(* IEC 61131-3 sources: 2026_Projet_YGO_ExcavatriceDragage/TOOLS/TEST_AUTO_CI/RESULTS/L_SIMULATION/tests (part 9) *)

TEST 'TC-T418-INT-007 Config maintien reel trop long refuse sans bypass'
nx := 5000; ny := 5000; raw1 := 0; raw2 := 0; previousButton := FALSE; buttonEdges := 0;
bench.Enable := TRUE; joy.Enable := TRUE; joy.ArmingPermit := TRUE; diagOk.Operational := TRUE;
joy.BusCanOpenOP := diagOk; joy.JoystickOP := diagOk; home.Enable := TRUE; home.BootReady := TRUE;
home.Mode := E_Mode.MAINT_N1; home.BucketOffsetValid := TRUE; home.WinchesMechanicallyStopped := TRUE;
cfg.DeadmanArmHoldTime := T#1S;
ADVANCE_TIME(10000000);
bench(RawPosM1 := raw1, RawPosM2 := raw2);
joy(RawX := bench.Operator.JoyXRaw_ANA1, RawY := bench.Operator.JoyYRaw_ANA2, RawButton := bench.Operator.JoyBtnRaw, Cfg := cfg, NeutralXMem := nx, NeutralYMem := ny);
home(DeadmanArmed := joy.DeadmanArmed, JoystickDeflected := NOT joy.AtNeutralXY, JoystickPull := joy.AxisCmdY.DirectionPositive, JoystickPush := joy.AxisCmdY.DirectionNegative, BtnValidation := bench.Operator.JoyBtnRaw);
IF bench.Operator.JoyBtnRaw AND NOT previousButton THEN buttonEdges := buttonEdges + 1; END_IF; previousButton := bench.Operator.JoyBtnRaw;
bench.SimJoystickRight_Fwd_MAINT_Active := TRUE;
ADVANCE_TIME(10000000);
bench(RawPosM1 := raw1, RawPosM2 := raw2);
joy(RawX := bench.Operator.JoyXRaw_ANA1, RawY := bench.Operator.JoyYRaw_ANA2, RawButton := bench.Operator.JoyBtnRaw, Cfg := cfg, NeutralXMem := nx, NeutralYMem := ny);
home(DeadmanArmed := joy.DeadmanArmed, JoystickDeflected := NOT joy.AtNeutralXY, JoystickPull := joy.AxisCmdY.DirectionPositive, JoystickPush := joy.AxisCmdY.DirectionNegative, BtnValidation := bench.Operator.JoyBtnRaw);
IF bench.Operator.JoyBtnRaw AND NOT previousButton THEN buttonEdges := buttonEdges + 1; END_IF; previousButton := bench.Operator.JoyBtnRaw;
ASSERT_FALSE(joy.DeadmanArmed, 'Maintien reel superieur a appui simule donc refus'); ASSERT_FALSE(joy.AxisCmdX.StartStop, 'Aucun bypass');
ADVANCE_TIME(10000000);
bench(RawPosM1 := raw1, RawPosM2 := raw2);
joy(RawX := bench.Operator.JoyXRaw_ANA1, RawY := bench.Operator.JoyYRaw_ANA2, RawButton := bench.Operator.JoyBtnRaw, Cfg := cfg, NeutralXMem := nx, NeutralYMem := ny);
home(DeadmanArmed := joy.DeadmanArmed, JoystickDeflected := NOT joy.AtNeutralXY, JoystickPull := joy.AxisCmdY.DirectionPositive, JoystickPush := joy.AxisCmdY.DirectionNegative, BtnValidation := bench.Operator.JoyBtnRaw);
IF bench.Operator.JoyBtnRaw AND NOT previousButton THEN buttonEdges := buttonEdges + 1; END_IF; previousButton := bench.Operator.JoyBtnRaw;
ASSERT_FALSE(joy.DeadmanArmed, 'Maintien reel superieur a appui simule donc refus'); ASSERT_FALSE(joy.AxisCmdX.StartStop, 'Aucun bypass');
ADVANCE_TIME(10000000);
bench(RawPosM1 := raw1, RawPosM2 := raw2);
joy(RawX := bench.Operator.JoyXRaw_ANA1, RawY := bench.Operator.JoyYRaw_ANA2, RawButton := bench.Operator.JoyBtnRaw, Cfg := cfg, NeutralXMem := nx, NeutralYMem := ny);
home(DeadmanArmed := joy.DeadmanArmed, JoystickDeflected := NOT joy.AtNeutralXY, JoystickPull := joy.AxisCmdY.DirectionPositive, JoystickPush := joy.AxisCmdY.DirectionNegative, BtnValidation := bench.Operator.JoyBtnRaw);
IF bench.Operator.JoyBtnRaw AND NOT previousButton THEN buttonEdges := buttonEdges + 1; END_IF; previousButton := bench.Operator.JoyBtnRaw;
ASSERT_FALSE(joy.DeadmanArmed, 'Maintien reel superieur a appui simule donc refus'); ASSERT_FALSE(joy.AxisCmdX.StartStop, 'Aucun bypass');
ADVANCE_TIME(10000000);
bench(RawPosM1 := raw1, RawPosM2 := raw2);
joy(RawX := bench.Operator.JoyXRaw_ANA1, RawY := bench.Operator.JoyYRaw_ANA2, RawButton := bench.Operator.JoyBtnRaw, Cfg := cfg, NeutralXMem := nx, NeutralYMem := ny);
home(DeadmanArmed := joy.DeadmanArmed, JoystickDeflected := NOT joy.AtNeutralXY, JoystickPull := joy.AxisCmdY.DirectionPositive, JoystickPush := joy.AxisCmdY.DirectionNegative, BtnValidation := bench.Operator.JoyBtnRaw);
IF bench.Operator.JoyBtnRaw AND NOT previousButton THEN buttonEdges := buttonEdges + 1; END_IF; previousButton := bench.Operator.JoyBtnRaw;
ASSERT_FALSE(joy.DeadmanArmed, 'Maintien reel superieur a appui simule donc refus'); ASSERT_FALSE(joy.AxisCmdX.StartStop, 'Aucun bypass');
ADVANCE_TIME(10000000);
bench(RawPosM1 := raw1, RawPosM2 := raw2);
joy(RawX := bench.Operator.JoyXRaw_ANA1, RawY := bench.Operator.JoyYRaw_ANA2, RawButton := bench.Operator.JoyBtnRaw, Cfg := cfg, NeutralXMem := nx, NeutralYMem := ny);
home(DeadmanArmed := joy.DeadmanArmed, JoystickDeflected := NOT joy.AtNeutralXY, JoystickPull := joy.AxisCmdY.DirectionPositive, JoystickPush := joy.AxisCmdY.DirectionNegative, BtnValidation := bench.Operator.JoyBtnRaw);
IF bench.Operator.JoyBtnRaw AND NOT previousButton THEN buttonEdges := buttonEdges + 1; END_IF; previousButton := bench.Operator.JoyBtnRaw;
ASSERT_FALSE(joy.DeadmanArmed, 'Maintien reel superieur a appui simule donc refus'); ASSERT_FALSE(joy.AxisCmdX.StartStop, 'Aucun bypass');
ADVANCE_TIME(10000000);
bench(RawPosM1 := raw1, RawPosM2 := raw2);
joy(RawX := bench.Operator.JoyXRaw_ANA1, RawY := bench.Operator.JoyYRaw_ANA2, RawButton := bench.Operator.JoyBtnRaw, Cfg := cfg, NeutralXMem := nx, NeutralYMem := ny);
home(DeadmanArmed := joy.DeadmanArmed, JoystickDeflected := NOT joy.AtNeutralXY, JoystickPull := joy.AxisCmdY.DirectionPositive, JoystickPush := joy.AxisCmdY.DirectionNegative, BtnValidation := bench.Operator.JoyBtnRaw);
IF bench.Operator.JoyBtnRaw AND NOT previousButton THEN buttonEdges := buttonEdges + 1; END_IF; previousButton := bench.Operator.JoyBtnRaw;
ASSERT_FALSE(joy.DeadmanArmed, 'Maintien reel superieur a appui simule donc refus'); ASSERT_FALSE(joy.AxisCmdX.StartStop, 'Aucun bypass');
ADVANCE_TIME(10000000);
bench(RawPosM1 := raw1, RawPosM2 := raw2);
joy(RawX := bench.Operator.JoyXRaw_ANA1, RawY := bench.Operator.JoyYRaw_ANA2, RawButton := bench.Operator.JoyBtnRaw, Cfg := cfg, NeutralXMem := nx, NeutralYMem := ny);
home(DeadmanArmed := joy.DeadmanArmed, JoystickDeflected := NOT joy.AtNeutralXY, JoystickPull := joy.AxisCmdY.DirectionPositive, JoystickPush := joy.AxisCmdY.DirectionNegative, BtnValidation := bench.Operator.JoyBtnRaw);
IF bench.Operator.JoyBtnRaw AND NOT previousButton THEN buttonEdges := buttonEdges + 1; END_IF; previousButton := bench.Operator.JoyBtnRaw;
ASSERT_FALSE(joy.DeadmanArmed, 'Maintien reel superieur a appui simule donc refus'); ASSERT_FALSE(joy.AxisCmdX.StartStop, 'Aucun bypass');
ADVANCE_TIME(10000000);
bench(RawPosM1 := raw1, RawPosM2 := raw2);
joy(RawX := bench.Operator.JoyXRaw_ANA1, RawY := bench.Operator.JoyYRaw_ANA2, RawButton := bench.Operator.JoyBtnRaw, Cfg := cfg, NeutralXMem := nx, NeutralYMem := ny);
home(DeadmanArmed := joy.DeadmanArmed, JoystickDeflected := NOT joy.AtNeutralXY, JoystickPull := joy.AxisCmdY.DirectionPositive, JoystickPush := joy.AxisCmdY.DirectionNegative, BtnValidation := bench.Operator.JoyBtnRaw);
IF bench.Operator.JoyBtnRaw AND NOT previousButton THEN buttonEdges := buttonEdges + 1; END_IF; previousButton := bench.Operator.JoyBtnRaw;
ASSERT_FALSE(joy.DeadmanArmed, 'Maintien reel superieur a appui simule donc refus'); ASSERT_FALSE(joy.AxisCmdX.StartStop, 'Aucun bypass');
ADVANCE_TIME(10000000);
bench(RawPosM1 := raw1, RawPosM2 := raw2);
joy(RawX := bench.Operator.JoyXRaw_ANA1, RawY := bench.Operator.JoyYRaw_ANA2, RawButton := bench.Operator.JoyBtnRaw, Cfg := cfg, NeutralXMem := nx, NeutralYMem := ny);
home(DeadmanArmed := joy.DeadmanArmed, JoystickDeflected := NOT joy.AtNeutralXY, JoystickPull := joy.AxisCmdY.DirectionPositive, JoystickPush := joy.AxisCmdY.DirectionNegative, BtnValidation := bench.Operator.JoyBtnRaw);
IF bench.Operator.JoyBtnRaw AND NOT previousButton THEN buttonEdges := buttonEdges + 1; END_IF; previousButton := bench.Operator.JoyBtnRaw;
ASSERT_FALSE(joy.DeadmanArmed, 'Maintien reel superieur a appui simule donc refus'); ASSERT_FALSE(joy.AxisCmdX.StartStop, 'Aucun bypass');
ADVANCE_TIME(10000000);
bench(RawPosM1 := raw1, RawPosM2 := raw2);
joy(RawX := bench.Operator.JoyXRaw_ANA1, RawY := bench.Operator.JoyYRaw_ANA2, RawButton := bench.Operator.JoyBtnRaw, Cfg := cfg, NeutralXMem := nx, NeutralYMem := ny);
home(DeadmanArmed := joy.DeadmanArmed, JoystickDeflected := NOT joy.AtNeutralXY, JoystickPull := joy.AxisCmdY.DirectionPositive, JoystickPush := joy.AxisCmdY.DirectionNegative, BtnValidation := bench.Operator.JoyBtnRaw);
IF bench.Operator.JoyBtnRaw AND NOT previousButton THEN buttonEdges := buttonEdges + 1; END_IF; previousButton := bench.Operator.JoyBtnRaw;
ASSERT_FALSE(joy.DeadmanArmed, 'Maintien reel superieur a appui simule donc refus'); ASSERT_FALSE(joy.AxisCmdX.StartStop, 'Aucun bypass');
ADVANCE_TIME(10000000);
bench(RawPosM1 := raw1, RawPosM2 := raw2);
joy(RawX := bench.Operator.JoyXRaw_ANA1, RawY := bench.Operator.JoyYRaw_ANA2, RawButton := bench.Operator.JoyBtnRaw, Cfg := cfg, NeutralXMem := nx, NeutralYMem := ny);
home(DeadmanArmed := joy.DeadmanArmed, JoystickDeflected := NOT joy.AtNeutralXY, JoystickPull := joy.AxisCmdY.DirectionPositive, JoystickPush := joy.AxisCmdY.DirectionNegative, BtnValidation := bench.Operator.JoyBtnRaw);
IF bench.Operator.JoyBtnRaw AND NOT previousButton THEN buttonEdges := buttonEdges + 1; END_IF; previousButton := bench.Operator.JoyBtnRaw;
ASSERT_FALSE(joy.DeadmanArmed, 'Maintien reel superieur a appui simule donc refus'); ASSERT_FALSE(joy.AxisCmdX.StartStop, 'Aucun bypass');
ADVANCE_TIME(10000000);
bench(RawPosM1 := raw1, RawPosM2 := raw2);
joy(RawX := bench.Operator.JoyXRaw_ANA1, RawY := bench.Operator.JoyYRaw_ANA2, RawButton := bench.Operator.JoyBtnRaw, Cfg := cfg, NeutralXMem := nx, NeutralYMem := ny);
home(DeadmanArmed := joy.DeadmanArmed, JoystickDeflected := NOT joy.AtNeutralXY, JoystickPull := joy.AxisCmdY.DirectionPositive, JoystickPush := joy.AxisCmdY.DirectionNegative, BtnValidation := bench.Operator.JoyBtnRaw);
IF bench.Operator.JoyBtnRaw AND NOT previousButton THEN buttonEdges := buttonEdges + 1; END_IF; previousButton := bench.Operator.JoyBtnRaw;
ASSERT_FALSE(joy.DeadmanArmed, 'Maintien reel superieur a appui simule donc refus'); ASSERT_FALSE(joy.AxisCmdX.StartStop, 'Aucun bypass');
ADVANCE_TIME(10000000);
bench(RawPosM1 := raw1, RawPosM2 := raw2);
joy(RawX := bench.Operator.JoyXRaw_ANA1, RawY := bench.Operator.JoyYRaw_ANA2, RawButton := bench.Operator.JoyBtnRaw, Cfg := cfg, NeutralXMem := nx, NeutralYMem := ny);
home(DeadmanArmed := joy.DeadmanArmed, JoystickDeflected := NOT joy.AtNeutralXY, JoystickPull := joy.AxisCmdY.DirectionPositive, JoystickPush := joy.AxisCmdY.DirectionNegative, BtnValidation := bench.Operator.JoyBtnRaw);
IF bench.Operator.JoyBtnRaw AND NOT previousButton THEN buttonEdges := buttonEdges + 1; END_IF; previousButton := bench.Operator.JoyBtnRaw;
ASSERT_FALSE(joy.DeadmanArmed, 'Maintien reel superieur a appui simule donc refus'); ASSERT_FALSE(joy.AxisCmdX.StartStop, 'Aucun bypass');
ADVANCE_TIME(10000000);
bench(RawPosM1 := raw1, RawPosM2 := raw2);
joy(RawX := bench.Operator.JoyXRaw_ANA1, RawY := bench.Operator.JoyYRaw_ANA2, RawButton := bench.Operator.JoyBtnRaw, Cfg := cfg, NeutralXMem := nx, NeutralYMem := ny);
home(DeadmanArmed := joy.DeadmanArmed, JoystickDeflected := NOT joy.AtNeutralXY, JoystickPull := joy.AxisCmdY.DirectionPositive, JoystickPush := joy.AxisCmdY.DirectionNegative, BtnValidation := bench.Operator.JoyBtnRaw);
IF bench.Operator.JoyBtnRaw AND NOT previousButton THEN buttonEdges := buttonEdges + 1; END_IF; previousButton := bench.Operator.JoyBtnRaw;
ASSERT_FALSE(joy.DeadmanArmed, 'Maintien reel superieur a appui simule donc refus'); ASSERT_FALSE(joy.AxisCmdX.StartStop, 'Aucun bypass');
ADVANCE_TIME(10000000);
bench(RawPosM1 := raw1, RawPosM2 := raw2);
joy(RawX := bench.Operator.JoyXRaw_ANA1, RawY := bench.Operator.JoyYRaw_ANA2, RawButton := bench.Operator.JoyBtnRaw, Cfg := cfg, NeutralXMem := nx, NeutralYMem := ny);
home(DeadmanArmed := joy.DeadmanArmed, JoystickDeflected := NOT joy.AtNeutralXY, JoystickPull := joy.AxisCmdY.DirectionPositive, JoystickPush := joy.AxisCmdY.DirectionNegative, BtnValidation := bench.Operator.JoyBtnRaw);
IF bench.Operator.JoyBtnRaw AND NOT previousButton THEN buttonEdges := buttonEdges + 1; END_IF; previousButton := bench.Operator.JoyBtnRaw;
ASSERT_FALSE(joy.DeadmanArmed, 'Maintien reel superieur a appui simule donc refus'); ASSERT_FALSE(joy.AxisCmdX.StartStop, 'Aucun bypass');
ADVANCE_TIME(10000000);
bench(RawPosM1 := raw1, RawPosM2 := raw2);
joy(RawX := bench.Operator.JoyXRaw_ANA1, RawY := bench.Operator.JoyYRaw_ANA2, RawButton := bench.Operator.JoyBtnRaw, Cfg := cfg, NeutralXMem := nx, NeutralYMem := ny);
home(DeadmanArmed := joy.DeadmanArmed, JoystickDeflected := NOT joy.AtNeutralXY, JoystickPull := joy.AxisCmdY.DirectionPositive, JoystickPush := joy.AxisCmdY.DirectionNegative, BtnValidation := bench.Operator.JoyBtnRaw);
IF bench.Operator.JoyBtnRaw AND NOT previousButton THEN buttonEdges := buttonEdges + 1; END_IF; previousButton := bench.Operator.JoyBtnRaw;
ASSERT_FALSE(joy.DeadmanArmed, 'Maintien reel superieur a appui simule donc refus'); ASSERT_FALSE(joy.AxisCmdX.StartStop, 'Aucun bypass');
ADVANCE_TIME(10000000);
bench(RawPosM1 := raw1, RawPosM2 := raw2);
joy(RawX := bench.Operator.JoyXRaw_ANA1, RawY := bench.Operator.JoyYRaw_ANA2, RawButton := bench.Operator.JoyBtnRaw, Cfg := cfg, NeutralXMem := nx, NeutralYMem := ny);
home(DeadmanArmed := joy.DeadmanArmed, JoystickDeflected := NOT joy.AtNeutralXY, JoystickPull := joy.AxisCmdY.DirectionPositive, JoystickPush := joy.AxisCmdY.DirectionNegative, BtnValidation := bench.Operator.JoyBtnRaw);
IF bench.Operator.JoyBtnRaw AND NOT previousButton THEN buttonEdges := buttonEdges + 1; END_IF; previousButton := bench.Operator.JoyBtnRaw;
ASSERT_FALSE(joy.DeadmanArmed, 'Maintien reel superieur a appui simule donc refus'); ASSERT_FALSE(joy.AxisCmdX.StartStop, 'Aucun bypass');
ADVANCE_TIME(10000000);
bench(RawPosM1 := raw1, RawPosM2 := raw2);
joy(RawX := bench.Operator.JoyXRaw_ANA1, RawY := bench.Operator.JoyYRaw_ANA2, RawButton := bench.Operator.JoyBtnRaw, Cfg := cfg, NeutralXMem := nx, NeutralYMem := ny);
home(DeadmanArmed := joy.DeadmanArmed, JoystickDeflected := NOT joy.AtNeutralXY, JoystickPull := joy.AxisCmdY.DirectionPositive, JoystickPush := joy.AxisCmdY.DirectionNegative, BtnValidation := bench.Operator.JoyBtnRaw);
IF bench.Operator.JoyBtnRaw AND NOT previousButton THEN buttonEdges := buttonEdges + 1; END_IF; previousButton := bench.Operator.JoyBtnRaw;
ASSERT_FALSE(joy.DeadmanArmed, 'Maintien reel superieur a appui simule donc refus'); ASSERT_FALSE(joy.AxisCmdX.StartStop, 'Aucun bypass');
ADVANCE_TIME(10000000);
bench(RawPosM1 := raw1, RawPosM2 := raw2);
joy(RawX := bench.Operator.JoyXRaw_ANA1, RawY := bench.Operator.JoyYRaw_ANA2, RawButton := bench.Operator.JoyBtnRaw, Cfg := cfg, NeutralXMem := nx, NeutralYMem := ny);
home(DeadmanArmed := joy.DeadmanArmed, JoystickDeflected := NOT joy.AtNeutralXY, JoystickPull := joy.AxisCmdY.DirectionPositive, JoystickPush := joy.AxisCmdY.DirectionNegative, BtnValidation := bench.Operator.JoyBtnRaw);
IF bench.Operator.JoyBtnRaw AND NOT previousButton THEN buttonEdges := buttonEdges + 1; END_IF; previousButton := bench.Operator.JoyBtnRaw;
ASSERT_FALSE(joy.DeadmanArmed, 'Maintien reel superieur a appui simule donc refus'); ASSERT_FALSE(joy.AxisCmdX.StartStop, 'Aucun bypass');
ADVANCE_TIME(10000000);
bench(RawPosM1 := raw1, RawPosM2 := raw2);
joy(RawX := bench.Operator.JoyXRaw_ANA1, RawY := bench.Operator.JoyYRaw_ANA2, RawButton := bench.Operator.JoyBtnRaw, Cfg := cfg, NeutralXMem := nx, NeutralYMem := ny);
home(DeadmanArmed := joy.DeadmanArmed, JoystickDeflected := NOT joy.AtNeutralXY, JoystickPull := joy.AxisCmdY.DirectionPositive, JoystickPush := joy.AxisCmdY.DirectionNegative, BtnValidation := bench.Operator.JoyBtnRaw);
IF bench.Operator.JoyBtnRaw AND NOT previousButton THEN buttonEdges := buttonEdges + 1; END_IF; previousButton := bench.Operator.JoyBtnRaw;
ASSERT_FALSE(joy.DeadmanArmed, 'Maintien reel superieur a appui simule donc refus'); ASSERT_FALSE(joy.AxisCmdX.StartStop, 'Aucun bypass');
ADVANCE_TIME(10000000);
bench(RawPosM1 := raw1, RawPosM2 := raw2);
joy(RawX := bench.Operator.JoyXRaw_ANA1, RawY := bench.Operator.JoyYRaw_ANA2, RawButton := bench.Operator.JoyBtnRaw, Cfg := cfg, NeutralXMem := nx, NeutralYMem := ny);
home(DeadmanArmed := joy.DeadmanArmed, JoystickDeflected := NOT joy.AtNeutralXY, JoystickPull := joy.AxisCmdY.DirectionPositive, JoystickPush := joy.AxisCmdY.DirectionNegative, BtnValidation := bench.Operator.JoyBtnRaw);
IF bench.Operator.JoyBtnRaw AND NOT previousButton THEN buttonEdges := buttonEdges + 1; END_IF; previousButton := bench.Operator.JoyBtnRaw;
ASSERT_FALSE(joy.DeadmanArmed, 'Maintien reel superieur a appui simule donc refus'); ASSERT_FALSE(joy.AxisCmdX.StartStop, 'Aucun bypass');
ADVANCE_TIME(10000000);
bench(RawPosM1 := raw1, RawPosM2 := raw2);
joy(RawX := bench.Operator.JoyXRaw_ANA1, RawY := bench.Operator.JoyYRaw_ANA2, RawButton := bench.Operator.JoyBtnRaw, Cfg := cfg, NeutralXMem := nx, NeutralYMem := ny);
home(DeadmanArmed := joy.DeadmanArmed, JoystickDeflected := NOT joy.AtNeutralXY, JoystickPull := joy.AxisCmdY.DirectionPositive, JoystickPush := joy.AxisCmdY.DirectionNegative, BtnValidation := bench.Operator.JoyBtnRaw);
IF bench.Operator.JoyBtnRaw AND NOT previousButton THEN buttonEdges := buttonEdges + 1; END_IF; previousButton := bench.Operator.JoyBtnRaw;
ASSERT_FALSE(joy.DeadmanArmed, 'Maintien reel superieur a appui simule donc refus'); ASSERT_FALSE(joy.AxisCmdX.StartStop, 'Aucun bypass');
ADVANCE_TIME(10000000);
bench(RawPosM1 := raw1, RawPosM2 := raw2);
joy(RawX := bench.Operator.JoyXRaw_ANA1, RawY := bench.Operator.JoyYRaw_ANA2, RawButton := bench.Operator.JoyBtnRaw, Cfg := cfg, NeutralXMem := nx, NeutralYMem := ny);
home(DeadmanArmed := joy.DeadmanArmed, JoystickDeflected := NOT joy.AtNeutralXY, JoystickPull := joy.AxisCmdY.DirectionPositive, JoystickPush := joy.AxisCmdY.DirectionNegative, BtnValidation := bench.Operator.JoyBtnRaw);
IF bench.Operator.JoyBtnRaw AND NOT previousButton THEN buttonEdges := buttonEdges + 1; END_IF; previousButton := bench.Operator.JoyBtnRaw;
ASSERT_FALSE(joy.DeadmanArmed, 'Maintien reel superieur a appui simule donc refus'); ASSERT_FALSE(joy.AxisCmdX.StartStop, 'Aucun bypass');
ADVANCE_TIME(10000000);
bench(RawPosM1 := raw1, RawPosM2 := raw2);
joy(RawX := bench.Operator.JoyXRaw_ANA1, RawY := bench.Operator.JoyYRaw_ANA2, RawButton := bench.Operator.JoyBtnRaw, Cfg := cfg, NeutralXMem := nx, NeutralYMem := ny);
home(DeadmanArmed := joy.DeadmanArmed, JoystickDeflected := NOT joy.AtNeutralXY, JoystickPull := joy.AxisCmdY.DirectionPositive, JoystickPush := joy.AxisCmdY.DirectionNegative, BtnValidation := bench.Operator.JoyBtnRaw);
IF bench.Operator.JoyBtnRaw AND NOT previousButton THEN buttonEdges := buttonEdges + 1; END_IF; previousButton := bench.Operator.JoyBtnRaw;
ASSERT_FALSE(joy.DeadmanArmed, 'Maintien reel superieur a appui simule donc refus'); ASSERT_FALSE(joy.AxisCmdX.StartStop, 'Aucun bypass');
ADVANCE_TIME(10000000);
bench(RawPosM1 := raw1, RawPosM2 := raw2);
joy(RawX := bench.Operator.JoyXRaw_ANA1, RawY := bench.Operator.JoyYRaw_ANA2, RawButton := bench.Operator.JoyBtnRaw, Cfg := cfg, NeutralXMem := nx, NeutralYMem := ny);
home(DeadmanArmed := joy.DeadmanArmed, JoystickDeflected := NOT joy.AtNeutralXY, JoystickPull := joy.AxisCmdY.DirectionPositive, JoystickPush := joy.AxisCmdY.DirectionNegative, BtnValidation := bench.Operator.JoyBtnRaw);
IF bench.Operator.JoyBtnRaw AND NOT previousButton THEN buttonEdges := buttonEdges + 1; END_IF; previousButton := bench.Operator.JoyBtnRaw;
ASSERT_FALSE(joy.DeadmanArmed, 'Maintien reel superieur a appui simule donc refus'); ASSERT_FALSE(joy.AxisCmdX.StartStop, 'Aucun bypass');
ADVANCE_TIME(10000000);
bench(RawPosM1 := raw1, RawPosM2 := raw2);
joy(RawX := bench.Operator.JoyXRaw_ANA1, RawY := bench.Operator.JoyYRaw_ANA2, RawButton := bench.Operator.JoyBtnRaw, Cfg := cfg, NeutralXMem := nx, NeutralYMem := ny);
home(DeadmanArmed := joy.DeadmanArmed, JoystickDeflected := NOT joy.AtNeutralXY, JoystickPull := joy.AxisCmdY.DirectionPositive, JoystickPush := joy.AxisCmdY.DirectionNegative, BtnValidation := bench.Operator.JoyBtnRaw);
IF bench.Operator.JoyBtnRaw AND NOT previousButton THEN buttonEdges := buttonEdges + 1; END_IF; previousButton := bench.Operator.JoyBtnRaw;
ASSERT_FALSE(joy.DeadmanArmed, 'Maintien reel superieur a appui simule donc refus'); ASSERT_FALSE(joy.AxisCmdX.StartStop, 'Aucun bypass');
ADVANCE_TIME(10000000);
bench(RawPosM1 := raw1, RawPosM2 := raw2);
joy(RawX := bench.Operator.JoyXRaw_ANA1, RawY := bench.Operator.JoyYRaw_ANA2, RawButton := bench.Operator.JoyBtnRaw, Cfg := cfg, NeutralXMem := nx, NeutralYMem := ny);
home(DeadmanArmed := joy.DeadmanArmed, JoystickDeflected := NOT joy.AtNeutralXY, JoystickPull := joy.AxisCmdY.DirectionPositive, JoystickPush := joy.AxisCmdY.DirectionNegative, BtnValidation := bench.Operator.JoyBtnRaw);
IF bench.Operator.JoyBtnRaw AND NOT previousButton THEN buttonEdges := buttonEdges + 1; END_IF; previousButton := bench.Operator.JoyBtnRaw;
ASSERT_FALSE(joy.DeadmanArmed, 'Maintien reel superieur a appui simule donc refus'); ASSERT_FALSE(joy.AxisCmdX.StartStop, 'Aucun bypass');
ADVANCE_TIME(10000000);
bench(RawPosM1 := raw1, RawPosM2 := raw2);
joy(RawX := bench.Operator.JoyXRaw_ANA1, RawY := bench.Operator.JoyYRaw_ANA2, RawButton := bench.Operator.JoyBtnRaw, Cfg := cfg, NeutralXMem := nx, NeutralYMem := ny);
home(DeadmanArmed := joy.DeadmanArmed, JoystickDeflected := NOT joy.AtNeutralXY, JoystickPull := joy.AxisCmdY.DirectionPositive, JoystickPush := joy.AxisCmdY.DirectionNegative, BtnValidation := bench.Operator.JoyBtnRaw);
IF bench.Operator.JoyBtnRaw AND NOT previousButton THEN buttonEdges := buttonEdges + 1; END_IF; previousButton := bench.Operator.JoyBtnRaw;
ASSERT_FALSE(joy.DeadmanArmed, 'Maintien reel superieur a appui simule donc refus'); ASSERT_FALSE(joy.AxisCmdX.StartStop, 'Aucun bypass');
ADVANCE_TIME(10000000);
bench(RawPosM1 := raw1, RawPosM2 := raw2);
joy(RawX := bench.Operator.JoyXRaw_ANA1, RawY := bench.Operator.JoyYRaw_ANA2, RawButton := bench.Operator.JoyBtnRaw, Cfg := cfg, NeutralXMem := nx, NeutralYMem := ny);
home(DeadmanArmed := joy.DeadmanArmed, JoystickDeflected := NOT joy.AtNeutralXY, JoystickPull := joy.AxisCmdY.DirectionPositive, JoystickPush := joy.AxisCmdY.DirectionNegative, BtnValidation := bench.Operator.JoyBtnRaw);
IF bench.Operator.JoyBtnRaw AND NOT previousButton THEN buttonEdges := buttonEdges + 1; END_IF; previousButton := bench.Operator.JoyBtnRaw;
ASSERT_FALSE(joy.DeadmanArmed, 'Maintien reel superieur a appui simule donc refus'); ASSERT_FALSE(joy.AxisCmdX.StartStop, 'Aucun bypass');
ADVANCE_TIME(10000000);
bench(RawPosM1 := raw1, RawPosM2 := raw2);
joy(RawX := bench.Operator.JoyXRaw_ANA1, RawY := bench.Operator.JoyYRaw_ANA2, RawButton := bench.Operator.JoyBtnRaw, Cfg := cfg, NeutralXMem := nx, NeutralYMem := ny);
home(DeadmanArmed := joy.DeadmanArmed, JoystickDeflected := NOT joy.AtNeutralXY, JoystickPull := joy.AxisCmdY.DirectionPositive, JoystickPush := joy.AxisCmdY.DirectionNegative, BtnValidation := bench.Operator.JoyBtnRaw);
IF bench.Operator.JoyBtnRaw AND NOT previousButton THEN buttonEdges := buttonEdges + 1; END_IF; previousButton := bench.Operator.JoyBtnRaw;
ASSERT_FALSE(joy.DeadmanArmed, 'Maintien reel superieur a appui simule donc refus'); ASSERT_FALSE(joy.AxisCmdX.StartStop, 'Aucun bypass');
ADVANCE_TIME(10000000);
bench(RawPosM1 := raw1, RawPosM2 := raw2);
joy(RawX := bench.Operator.JoyXRaw_ANA1, RawY := bench.Operator.JoyYRaw_ANA2, RawButton := bench.Operator.JoyBtnRaw, Cfg := cfg, NeutralXMem := nx, NeutralYMem := ny);
home(DeadmanArmed := joy.DeadmanArmed, JoystickDeflected := NOT joy.AtNeutralXY, JoystickPull := joy.AxisCmdY.DirectionPositive, JoystickPush := joy.AxisCmdY.DirectionNegative, BtnValidation := bench.Operator.JoyBtnRaw);
IF bench.Operator.JoyBtnRaw AND NOT previousButton THEN buttonEdges := buttonEdges + 1; END_IF; previousButton := bench.Operator.JoyBtnRaw;
ASSERT_FALSE(joy.DeadmanArmed, 'Maintien reel superieur a appui simule donc refus'); ASSERT_FALSE(joy.AxisCmdX.StartStop, 'Aucun bypass');
ADVANCE_TIME(10000000);
bench(RawPosM1 := raw1, RawPosM2 := raw2);
joy(RawX := bench.Operator.JoyXRaw_ANA1, RawY := bench.Operator.JoyYRaw_ANA2, RawButton := bench.Operator.JoyBtnRaw, Cfg := cfg, NeutralXMem := nx, NeutralYMem := ny);
home(DeadmanArmed := joy.DeadmanArmed, JoystickDeflected := NOT joy.AtNeutralXY, JoystickPull := joy.AxisCmdY.DirectionPositive, JoystickPush := joy.AxisCmdY.DirectionNegative, BtnValidation := bench.Operator.JoyBtnRaw);
IF bench.Operator.JoyBtnRaw AND NOT previousButton THEN buttonEdges := buttonEdges + 1; END_IF; previousButton := bench.Operator.JoyBtnRaw;
ASSERT_FALSE(joy.DeadmanArmed, 'Maintien reel superieur a appui simule donc refus'); ASSERT_FALSE(joy.AxisCmdX.StartStop, 'Aucun bypass');
ADVANCE_TIME(10000000);
bench(RawPosM1 := raw1, RawPosM2 := raw2);
joy(RawX := bench.Operator.JoyXRaw_ANA1, RawY := bench.Operator.JoyYRaw_ANA2, RawButton := bench.Operator.JoyBtnRaw, Cfg := cfg, NeutralXMem := nx, NeutralYMem := ny);
home(DeadmanArmed := joy.DeadmanArmed, JoystickDeflected := NOT joy.AtNeutralXY, JoystickPull := joy.AxisCmdY.DirectionPositive, JoystickPush := joy.AxisCmdY.DirectionNegative, BtnValidation := bench.Operator.JoyBtnRaw);
IF bench.Operator.JoyBtnRaw AND NOT previousButton THEN buttonEdges := buttonEdges + 1; END_IF; previousButton := bench.Operator.JoyBtnRaw;
ASSERT_FALSE(joy.DeadmanArmed, 'Maintien reel superieur a appui simule donc refus'); ASSERT_FALSE(joy.AxisCmdX.StartStop, 'Aucun bypass');
ADVANCE_TIME(10000000);
bench(RawPosM1 := raw1, RawPosM2 := raw2);
joy(RawX := bench.Operator.JoyXRaw_ANA1, RawY := bench.Operator.JoyYRaw_ANA2, RawButton := bench.Operator.JoyBtnRaw, Cfg := cfg, NeutralXMem := nx, NeutralYMem := ny);
home(DeadmanArmed := joy.DeadmanArmed, JoystickDeflected := NOT joy.AtNeutralXY, JoystickPull := joy.AxisCmdY.DirectionPositive, JoystickPush := joy.AxisCmdY.DirectionNegative, BtnValidation := bench.Operator.JoyBtnRaw);
IF bench.Operator.JoyBtnRaw AND NOT previousButton THEN buttonEdges := buttonEdges + 1; END_IF; previousButton := bench.Operator.JoyBtnRaw;
ASSERT_FALSE(joy.DeadmanArmed, 'Maintien reel superieur a appui simule donc refus'); ASSERT_FALSE(joy.AxisCmdX.StartStop, 'Aucun bypass');
ADVANCE_TIME(10000000);
bench(RawPosM1 := raw1, RawPosM2 := raw2);
joy(RawX := bench.Operator.JoyXRaw_ANA1, RawY := bench.Operator.JoyYRaw_ANA2, RawButton := bench.Operator.JoyBtnRaw, Cfg := cfg, NeutralXMem := nx, NeutralYMem := ny);
home(DeadmanArmed := joy.DeadmanArmed, JoystickDeflected := NOT joy.AtNeutralXY, JoystickPull := joy.AxisCmdY.DirectionPositive, JoystickPush := joy.AxisCmdY.DirectionNegative, BtnValidation := bench.Operator.JoyBtnRaw);
IF bench.Operator.JoyBtnRaw AND NOT previousButton THEN buttonEdges := buttonEdges + 1; END_IF; previousButton := bench.Operator.JoyBtnRaw;
ASSERT_FALSE(joy.DeadmanArmed, 'Maintien reel superieur a appui simule donc refus'); ASSERT_FALSE(joy.AxisCmdX.StartStop, 'Aucun bypass');
ADVANCE_TIME(10000000);
bench(RawPosM1 := raw1, RawPosM2 := raw2);
joy(RawX := bench.Operator.JoyXRaw_ANA1, RawY := bench.Operator.JoyYRaw_ANA2, RawButton := bench.Operator.JoyBtnRaw, Cfg := cfg, NeutralXMem := nx, NeutralYMem := ny);
home(DeadmanArmed := joy.DeadmanArmed, JoystickDeflected := NOT joy.AtNeutralXY, JoystickPull := joy.AxisCmdY.DirectionPositive, JoystickPush := joy.AxisCmdY.DirectionNegative, BtnValidation := bench.Operator.JoyBtnRaw);
IF bench.Operator.JoyBtnRaw AND NOT previousButton THEN buttonEdges := buttonEdges + 1; END_IF; previousButton := bench.Operator.JoyBtnRaw;
ASSERT_FALSE(joy.DeadmanArmed, 'Maintien reel superieur a appui simule donc refus'); ASSERT_FALSE(joy.AxisCmdX.StartStop, 'Aucun bypass');
ADVANCE_TIME(10000000);
bench(RawPosM1 := raw1, RawPosM2 := raw2);
joy(RawX := bench.Operator.JoyXRaw_ANA1, RawY := bench.Operator.JoyYRaw_ANA2, RawButton := bench.Operator.JoyBtnRaw, Cfg := cfg, NeutralXMem := nx, NeutralYMem := ny);
home(DeadmanArmed := joy.DeadmanArmed, JoystickDeflected := NOT joy.AtNeutralXY, JoystickPull := joy.AxisCmdY.DirectionPositive, JoystickPush := joy.AxisCmdY.DirectionNegative, BtnValidation := bench.Operator.JoyBtnRaw);
IF bench.Operator.JoyBtnRaw AND NOT previousButton THEN buttonEdges := buttonEdges + 1; END_IF; previousButton := bench.Operator.JoyBtnRaw;
ASSERT_FALSE(joy.DeadmanArmed, 'Maintien reel superieur a appui simule donc refus'); ASSERT_FALSE(joy.AxisCmdX.StartStop, 'Aucun bypass');
ADVANCE_TIME(10000000);
bench(RawPosM1 := raw1, RawPosM2 := raw2);
joy(RawX := bench.Operator.JoyXRaw_ANA1, RawY := bench.Operator.JoyYRaw_ANA2, RawButton := bench.Operator.JoyBtnRaw, Cfg := cfg, NeutralXMem := nx, NeutralYMem := ny);
home(DeadmanArmed := joy.DeadmanArmed, JoystickDeflected := NOT joy.AtNeutralXY, JoystickPull := joy.AxisCmdY.DirectionPositive, JoystickPush := joy.AxisCmdY.DirectionNegative, BtnValidation := bench.Operator.JoyBtnRaw);
IF bench.Operator.JoyBtnRaw AND NOT previousButton THEN buttonEdges := buttonEdges + 1; END_IF; previousButton := bench.Operator.JoyBtnRaw;
ASSERT_FALSE(joy.DeadmanArmed, 'Maintien reel superieur a appui simule donc refus'); ASSERT_FALSE(joy.AxisCmdX.StartStop, 'Aucun bypass');
ADVANCE_TIME(10000000);
bench(RawPosM1 := raw1, RawPosM2 := raw2);
joy(RawX := bench.Operator.JoyXRaw_ANA1, RawY := bench.Operator.JoyYRaw_ANA2, RawButton := bench.Operator.JoyBtnRaw, Cfg := cfg, NeutralXMem := nx, NeutralYMem := ny);
home(DeadmanArmed := joy.DeadmanArmed, JoystickDeflected := NOT joy.AtNeutralXY, JoystickPull := joy.AxisCmdY.DirectionPositive, JoystickPush := joy.AxisCmdY.DirectionNegative, BtnValidation := bench.Operator.JoyBtnRaw);
IF bench.Operator.JoyBtnRaw AND NOT previousButton THEN buttonEdges := buttonEdges + 1; END_IF; previousButton := bench.Operator.JoyBtnRaw;
ASSERT_FALSE(joy.DeadmanArmed, 'Maintien reel superieur a appui simule donc refus'); ASSERT_FALSE(joy.AxisCmdX.StartStop, 'Aucun bypass');
ADVANCE_TIME(10000000);
bench(RawPosM1 := raw1, RawPosM2 := raw2);
joy(RawX := bench.Operator.JoyXRaw_ANA1, RawY := bench.Operator.JoyYRaw_ANA2, RawButton := bench.Operator.JoyBtnRaw, Cfg := cfg, NeutralXMem := nx, NeutralYMem := ny);
home(DeadmanArmed := joy.DeadmanArmed, JoystickDeflected := NOT joy.AtNeutralXY, JoystickPull := joy.AxisCmdY.DirectionPositive, JoystickPush := joy.AxisCmdY.DirectionNegative, BtnValidation := bench.Operator.JoyBtnRaw);
IF bench.Operator.JoyBtnRaw AND NOT previousButton THEN buttonEdges := buttonEdges + 1; END_IF; previousButton := bench.Operator.JoyBtnRaw;
ASSERT_FALSE(joy.DeadmanArmed, 'Maintien reel superieur a appui simule donc refus'); ASSERT_FALSE(joy.AxisCmdX.StartStop, 'Aucun bypass');
ADVANCE_TIME(10000000);
bench(RawPosM1 := raw1, RawPosM2 := raw2);
joy(RawX := bench.Operator.JoyXRaw_ANA1, RawY := bench.Operator.JoyYRaw_ANA2, RawButton := bench.Operator.JoyBtnRaw, Cfg := cfg, NeutralXMem := nx, NeutralYMem := ny);
home(DeadmanArmed := joy.DeadmanArmed, JoystickDeflected := NOT joy.AtNeutralXY, JoystickPull := joy.AxisCmdY.DirectionPositive, JoystickPush := joy.AxisCmdY.DirectionNegative, BtnValidation := bench.Operator.JoyBtnRaw);
IF bench.Operator.JoyBtnRaw AND NOT previousButton THEN buttonEdges := buttonEdges + 1; END_IF; previousButton := bench.Operator.JoyBtnRaw;
ASSERT_FALSE(joy.DeadmanArmed, 'Maintien reel superieur a appui simule donc refus'); ASSERT_FALSE(joy.AxisCmdX.StartStop, 'Aucun bypass');
ADVANCE_TIME(10000000);
bench(RawPosM1 := raw1, RawPosM2 := raw2);
joy(RawX := bench.Operator.JoyXRaw_ANA1, RawY := bench.Operator.JoyYRaw_ANA2, RawButton := bench.Operator.JoyBtnRaw, Cfg := cfg, NeutralXMem := nx, NeutralYMem := ny);
home(DeadmanArmed := joy.DeadmanArmed, JoystickDeflected := NOT joy.AtNeutralXY, JoystickPull := joy.AxisCmdY.DirectionPositive, JoystickPush := joy.AxisCmdY.DirectionNegative, BtnValidation := bench.Operator.JoyBtnRaw);
IF bench.Operator.JoyBtnRaw AND NOT previousButton THEN buttonEdges := buttonEdges + 1; END_IF; previousButton := bench.Operator.JoyBtnRaw;
ASSERT_FALSE(joy.DeadmanArmed, 'Maintien reel superieur a appui simule donc refus'); ASSERT_FALSE(joy.AxisCmdX.StartStop, 'Aucun bypass');
ADVANCE_TIME(10000000);
bench(RawPosM1 := raw1, RawPosM2 := raw2);
joy(RawX := bench.Operator.JoyXRaw_ANA1, RawY := bench.Operator.JoyYRaw_ANA2, RawButton := bench.Operator.JoyBtnRaw, Cfg := cfg, NeutralXMem := nx, NeutralYMem := ny);
home(DeadmanArmed := joy.DeadmanArmed, JoystickDeflected := NOT joy.AtNeutralXY, JoystickPull := joy.AxisCmdY.DirectionPositive, JoystickPush := joy.AxisCmdY.DirectionNegative, BtnValidation := bench.Operator.JoyBtnRaw);
IF bench.Operator.JoyBtnRaw AND NOT previousButton THEN buttonEdges := buttonEdges + 1; END_IF; previousButton := bench.Operator.JoyBtnRaw;
ASSERT_FALSE(joy.DeadmanArmed, 'Maintien reel superieur a appui simule donc refus'); ASSERT_FALSE(joy.AxisCmdX.StartStop, 'Aucun bypass');
ADVANCE_TIME(10000000);
bench(RawPosM1 := raw1, RawPosM2 := raw2);
joy(RawX := bench.Operator.JoyXRaw_ANA1, RawY := bench.Operator.JoyYRaw_ANA2, RawButton := bench.Operator.JoyBtnRaw, Cfg := cfg, NeutralXMem := nx, NeutralYMem := ny);
home(DeadmanArmed := joy.DeadmanArmed, JoystickDeflected := NOT joy.AtNeutralXY, JoystickPull := joy.AxisCmdY.DirectionPositive, JoystickPush := joy.AxisCmdY.DirectionNegative, BtnValidation := bench.Operator.JoyBtnRaw);
IF bench.Operator.JoyBtnRaw AND NOT previousButton THEN buttonEdges := buttonEdges + 1; END_IF; previousButton := bench.Operator.JoyBtnRaw;
ASSERT_FALSE(joy.DeadmanArmed, 'Maintien reel superieur a appui simule donc refus'); ASSERT_FALSE(joy.AxisCmdX.StartStop, 'Aucun bypass');
ADVANCE_TIME(10000000);
bench(RawPosM1 := raw1, RawPosM2 := raw2);
joy(RawX := bench.Operator.JoyXRaw_ANA1, RawY := bench.Operator.JoyYRaw_ANA2, RawButton := bench.Operator.JoyBtnRaw, Cfg := cfg, NeutralXMem := nx, NeutralYMem := ny);
home(DeadmanArmed := joy.DeadmanArmed, JoystickDeflected := NOT joy.AtNeutralXY, JoystickPull := joy.AxisCmdY.DirectionPositive, JoystickPush := joy.AxisCmdY.DirectionNegative, BtnValidation := bench.Operator.JoyBtnRaw);
IF bench.Operator.JoyBtnRaw AND NOT previousButton THEN buttonEdges := buttonEdges + 1; END_IF; previousButton := bench.Operator.JoyBtnRaw;
ASSERT_FALSE(joy.DeadmanArmed, 'Maintien reel superieur a appui simule donc refus'); ASSERT_FALSE(joy.AxisCmdX.StartStop, 'Aucun bypass');
ADVANCE_TIME(10000000);
bench(RawPosM1 := raw1, RawPosM2 := raw2);
joy(RawX := bench.Operator.JoyXRaw_ANA1, RawY := bench.Operator.JoyYRaw_ANA2, RawButton := bench.Operator.JoyBtnRaw, Cfg := cfg, NeutralXMem := nx, NeutralYMem := ny);
home(DeadmanArmed := joy.DeadmanArmed, JoystickDeflected := NOT joy.AtNeutralXY, JoystickPull := joy.AxisCmdY.DirectionPositive, JoystickPush := joy.AxisCmdY.DirectionNegative, BtnValidation := bench.Operator.JoyBtnRaw);
IF bench.Operator.JoyBtnRaw AND NOT previousButton THEN buttonEdges := buttonEdges + 1; END_IF; previousButton := bench.Operator.JoyBtnRaw;
ASSERT_FALSE(joy.DeadmanArmed, 'Maintien reel superieur a appui simule donc refus'); ASSERT_FALSE(joy.AxisCmdX.StartStop, 'Aucun bypass');
ADVANCE_TIME(10000000);
bench(RawPosM1 := raw1, RawPosM2 := raw2);
joy(RawX := bench.Operator.JoyXRaw_ANA1, RawY := bench.Operator.JoyYRaw_ANA2, RawButton := bench.Operator.JoyBtnRaw, Cfg := cfg, NeutralXMem := nx, NeutralYMem := ny);
home(DeadmanArmed := joy.DeadmanArmed, JoystickDeflected := NOT joy.AtNeutralXY, JoystickPull := joy.AxisCmdY.DirectionPositive, JoystickPush := joy.AxisCmdY.DirectionNegative, BtnValidation := bench.Operator.JoyBtnRaw);
IF bench.Operator.JoyBtnRaw AND NOT previousButton THEN buttonEdges := buttonEdges + 1; END_IF; previousButton := bench.Operator.JoyBtnRaw;
ASSERT_FALSE(joy.DeadmanArmed, 'Maintien reel superieur a appui simule donc refus'); ASSERT_FALSE(joy.AxisCmdX.StartStop, 'Aucun bypass');
ADVANCE_TIME(10000000);
bench(RawPosM1 := raw1, RawPosM2 := raw2);
joy(RawX := bench.Operator.JoyXRaw_ANA1, RawY := bench.Operator.JoyYRaw_ANA2, RawButton := bench.Operator.JoyBtnRaw, Cfg := cfg, NeutralXMem := nx, NeutralYMem := ny);
home(DeadmanArmed := joy.DeadmanArmed, JoystickDeflected := NOT joy.AtNeutralXY, JoystickPull := joy.AxisCmdY.DirectionPositive, JoystickPush := joy.AxisCmdY.DirectionNegative, BtnValidation := bench.Operator.JoyBtnRaw);
IF bench.Operator.JoyBtnRaw AND NOT previousButton THEN buttonEdges := buttonEdges + 1; END_IF; previousButton := bench.Operator.JoyBtnRaw;
ASSERT_FALSE(joy.DeadmanArmed, 'Maintien reel superieur a appui simule donc refus'); ASSERT_FALSE(joy.AxisCmdX.StartStop, 'Aucun bypass');
ADVANCE_TIME(10000000);
bench(RawPosM1 := raw1, RawPosM2 := raw2);
joy(RawX := bench.Operator.JoyXRaw_ANA1, RawY := bench.Operator.JoyYRaw_ANA2, RawButton := bench.Operator.JoyBtnRaw, Cfg := cfg, NeutralXMem := nx, NeutralYMem := ny);
home(DeadmanArmed := joy.DeadmanArmed, JoystickDeflected := NOT joy.AtNeutralXY, JoystickPull := joy.AxisCmdY.DirectionPositive, JoystickPush := joy.AxisCmdY.DirectionNegative, BtnValidation := bench.Operator.JoyBtnRaw);
IF bench.Operator.JoyBtnRaw AND NOT previousButton THEN buttonEdges := buttonEdges + 1; END_IF; previousButton := bench.Operator.JoyBtnRaw;
ASSERT_FALSE(joy.DeadmanArmed, 'Maintien reel superieur a appui simule donc refus'); ASSERT_FALSE(joy.AxisCmdX.StartStop, 'Aucun bypass');
ADVANCE_TIME(10000000);
bench(RawPosM1 := raw1, RawPosM2 := raw2);
joy(RawX := bench.Operator.JoyXRaw_ANA1, RawY := bench.Operator.JoyYRaw_ANA2, RawButton := bench.Operator.JoyBtnRaw, Cfg := cfg, NeutralXMem := nx, NeutralYMem := ny);
home(DeadmanArmed := joy.DeadmanArmed, JoystickDeflected := NOT joy.AtNeutralXY, JoystickPull := joy.AxisCmdY.DirectionPositive, JoystickPush := joy.AxisCmdY.DirectionNegative, BtnValidation := bench.Operator.JoyBtnRaw);
IF bench.Operator.JoyBtnRaw AND NOT previousButton THEN buttonEdges := buttonEdges + 1; END_IF; previousButton := bench.Operator.JoyBtnRaw;
ASSERT_FALSE(joy.DeadmanArmed, 'Maintien reel superieur a appui simule donc refus'); ASSERT_FALSE(joy.AxisCmdX.StartStop, 'Aucun bypass');
ADVANCE_TIME(10000000);
bench(RawPosM1 := raw1, RawPosM2 := raw2);
joy(RawX := bench.Operator.JoyXRaw_ANA1, RawY := bench.Operator.JoyYRaw_ANA2, RawButton := bench.Operator.JoyBtnRaw, Cfg := cfg, NeutralXMem := nx, NeutralYMem := ny);
home(DeadmanArmed := joy.DeadmanArmed, JoystickDeflected := NOT joy.AtNeutralXY, JoystickPull := joy.AxisCmdY.DirectionPositive, JoystickPush := joy.AxisCmdY.DirectionNegative, BtnValidation := bench.Operator.JoyBtnRaw);
IF bench.Operator.JoyBtnRaw AND NOT previousButton THEN buttonEdges := buttonEdges + 1; END_IF; previousButton := bench.Operator.JoyBtnRaw;
ASSERT_FALSE(joy.DeadmanArmed, 'Maintien reel superieur a appui simule donc refus'); ASSERT_FALSE(joy.AxisCmdX.StartStop, 'Aucun bypass');
ADVANCE_TIME(10000000);
bench(RawPosM1 := raw1, RawPosM2 := raw2);
joy(RawX := bench.Operator.JoyXRaw_ANA1, RawY := bench.Operator.JoyYRaw_ANA2, RawButton := bench.Operator.JoyBtnRaw, Cfg := cfg, NeutralXMem := nx, NeutralYMem := ny);
home(DeadmanArmed := joy.DeadmanArmed, JoystickDeflected := NOT joy.AtNeutralXY, JoystickPull := joy.AxisCmdY.DirectionPositive, JoystickPush := joy.AxisCmdY.DirectionNegative, BtnValidation := bench.Operator.JoyBtnRaw);
IF bench.Operator.JoyBtnRaw AND NOT previousButton THEN buttonEdges := buttonEdges + 1; END_IF; previousButton := bench.Operator.JoyBtnRaw;
ASSERT_FALSE(joy.DeadmanArmed, 'Maintien reel superieur a appui simule donc refus'); ASSERT_FALSE(joy.AxisCmdX.StartStop, 'Aucun bypass');
ADVANCE_TIME(10000000);
bench(RawPosM1 := raw1, RawPosM2 := raw2);
joy(RawX := bench.Operator.JoyXRaw_ANA1, RawY := bench.Operator.JoyYRaw_ANA2, RawButton := bench.Operator.JoyBtnRaw, Cfg := cfg, NeutralXMem := nx, NeutralYMem := ny);
home(DeadmanArmed := joy.DeadmanArmed, JoystickDeflected := NOT joy.AtNeutralXY, JoystickPull := joy.AxisCmdY.DirectionPositive, JoystickPush := joy.AxisCmdY.DirectionNegative, BtnValidation := bench.Operator.JoyBtnRaw);
IF bench.Operator.JoyBtnRaw AND NOT previousButton THEN buttonEdges := buttonEdges + 1; END_IF; previousButton := bench.Operator.JoyBtnRaw;
ASSERT_FALSE(joy.DeadmanArmed, 'Maintien reel superieur a appui simule donc refus'); ASSERT_FALSE(joy.AxisCmdX.StartStop, 'Aucun bypass');
ADVANCE_TIME(10000000);
bench(RawPosM1 := raw1, RawPosM2 := raw2);
joy(RawX := bench.Operator.JoyXRaw_ANA1, RawY := bench.Operator.JoyYRaw_ANA2, RawButton := bench.Operator.JoyBtnRaw, Cfg := cfg, NeutralXMem := nx, NeutralYMem := ny);
home(DeadmanArmed := joy.DeadmanArmed, JoystickDeflected := NOT joy.AtNeutralXY, JoystickPull := joy.AxisCmdY.DirectionPositive, JoystickPush := joy.AxisCmdY.DirectionNegative, BtnValidation := bench.Operator.JoyBtnRaw);
IF bench.Operator.JoyBtnRaw AND NOT previousButton THEN buttonEdges := buttonEdges + 1; END_IF; previousButton := bench.Operator.JoyBtnRaw;
ASSERT_FALSE(joy.DeadmanArmed, 'Maintien reel superieur a appui simule donc refus'); ASSERT_FALSE(joy.AxisCmdX.StartStop, 'Aucun bypass');
ADVANCE_TIME(10000000);
bench(RawPosM1 := raw1, RawPosM2 := raw2);
joy(RawX := bench.Operator.JoyXRaw_ANA1, RawY := bench.Operator.JoyYRaw_ANA2, RawButton := bench.Operator.JoyBtnRaw, Cfg := cfg, NeutralXMem := nx, NeutralYMem := ny);
home(DeadmanArmed := joy.DeadmanArmed, JoystickDeflected := NOT joy.AtNeutralXY, JoystickPull := joy.AxisCmdY.DirectionPositive, JoystickPush := joy.AxisCmdY.DirectionNegative, BtnValidation := bench.Operator.JoyBtnRaw);
IF bench.Operator.JoyBtnRaw AND NOT previousButton THEN buttonEdges := buttonEdges + 1; END_IF; previousButton := bench.Operator.JoyBtnRaw;
ASSERT_FALSE(joy.DeadmanArmed, 'Maintien reel superieur a appui simule donc refus'); ASSERT_FALSE(joy.AxisCmdX.StartStop, 'Aucun bypass');
ADVANCE_TIME(10000000);
bench(RawPosM1 := raw1, RawPosM2 := raw2);
joy(RawX := bench.Operator.JoyXRaw_ANA1, RawY := bench.Operator.JoyYRaw_ANA2, RawButton := bench.Operator.JoyBtnRaw, Cfg := cfg, NeutralXMem := nx, NeutralYMem := ny);
home(DeadmanArmed := joy.DeadmanArmed, JoystickDeflected := NOT joy.AtNeutralXY, JoystickPull := joy.AxisCmdY.DirectionPositive, JoystickPush := joy.AxisCmdY.DirectionNegative, BtnValidation := bench.Operator.JoyBtnRaw);
IF bench.Operator.JoyBtnRaw AND NOT previousButton THEN buttonEdges := buttonEdges + 1; END_IF; previousButton := bench.Operator.JoyBtnRaw;
ASSERT_FALSE(joy.DeadmanArmed, 'Maintien reel superieur a appui simule donc refus'); ASSERT_FALSE(joy.AxisCmdX.StartStop, 'Aucun bypass');
ADVANCE_TIME(10000000);
bench(RawPosM1 := raw1, RawPosM2 := raw2);
joy(RawX := bench.Operator.JoyXRaw_ANA1, RawY := bench.Operator.JoyYRaw_ANA2, RawButton := bench.Operator.JoyBtnRaw, Cfg := cfg, NeutralXMem := nx, NeutralYMem := ny);
home(DeadmanArmed := joy.DeadmanArmed, JoystickDeflected := NOT joy.AtNeutralXY, JoystickPull := joy.AxisCmdY.DirectionPositive, JoystickPush := joy.AxisCmdY.DirectionNegative, BtnValidation := bench.Operator.JoyBtnRaw);
IF bench.Operator.JoyBtnRaw AND NOT previousButton THEN buttonEdges := buttonEdges + 1; END_IF; previousButton := bench.Operator.JoyBtnRaw;
ASSERT_FALSE(joy.DeadmanArmed, 'Maintien reel superieur a appui simule donc refus'); ASSERT_FALSE(joy.AxisCmdX.StartStop, 'Aucun bypass');
ADVANCE_TIME(10000000);
bench(RawPosM1 := raw1, RawPosM2 := raw2);
joy(RawX := bench.Operator.JoyXRaw_ANA1, RawY := bench.Operator.JoyYRaw_ANA2, RawButton := bench.Operator.JoyBtnRaw, Cfg := cfg, NeutralXMem := nx, NeutralYMem := ny);
home(DeadmanArmed := joy.DeadmanArmed, JoystickDeflected := NOT joy.AtNeutralXY, JoystickPull := joy.AxisCmdY.DirectionPositive, JoystickPush := joy.AxisCmdY.DirectionNegative, BtnValidation := bench.Operator.JoyBtnRaw);
IF bench.Operator.JoyBtnRaw AND NOT previousButton THEN buttonEdges := buttonEdges + 1; END_IF; previousButton := bench.Operator.JoyBtnRaw;
ASSERT_FALSE(joy.DeadmanArmed, 'Maintien reel superieur a appui simule donc refus'); ASSERT_FALSE(joy.AxisCmdX.StartStop, 'Aucun bypass');
ADVANCE_TIME(10000000);
bench(RawPosM1 := raw1, RawPosM2 := raw2);
joy(RawX := bench.Operator.JoyXRaw_ANA1, RawY := bench.Operator.JoyYRaw_ANA2, RawButton := bench.Operator.JoyBtnRaw, Cfg := cfg, NeutralXMem := nx, NeutralYMem := ny);
home(DeadmanArmed := joy.DeadmanArmed, JoystickDeflected := NOT joy.AtNeutralXY, JoystickPull := joy.AxisCmdY.DirectionPositive, JoystickPush := joy.AxisCmdY.DirectionNegative, BtnValidation := bench.Operator.JoyBtnRaw);
IF bench.Operator.JoyBtnRaw AND NOT previousButton THEN buttonEdges := buttonEdges + 1; END_IF; previousButton := bench.Operator.JoyBtnRaw;
ASSERT_FALSE(joy.DeadmanArmed, 'Maintien reel superieur a appui simule donc refus'); ASSERT_FALSE(joy.AxisCmdX.StartStop, 'Aucun bypass');
ADVANCE_TIME(10000000);
bench(RawPosM1 := raw1, RawPosM2 := raw2);
joy(RawX := bench.Operator.JoyXRaw_ANA1, RawY := bench.Operator.JoyYRaw_ANA2, RawButton := bench.Operator.JoyBtnRaw, Cfg := cfg, NeutralXMem := nx, NeutralYMem := ny);
home(DeadmanArmed := joy.DeadmanArmed, JoystickDeflected := NOT joy.AtNeutralXY, JoystickPull := joy.AxisCmdY.DirectionPositive, JoystickPush := joy.AxisCmdY.DirectionNegative, BtnValidation := bench.Operator.JoyBtnRaw);
IF bench.Operator.JoyBtnRaw AND NOT previousButton THEN buttonEdges := buttonEdges + 1; END_IF; previousButton := bench.Operator.JoyBtnRaw;
ASSERT_FALSE(joy.DeadmanArmed, 'Maintien reel superieur a appui simule donc refus'); ASSERT_FALSE(joy.AxisCmdX.StartStop, 'Aucun bypass');
ADVANCE_TIME(10000000);
bench(RawPosM1 := raw1, RawPosM2 := raw2);
joy(RawX := bench.Operator.JoyXRaw_ANA1, RawY := bench.Operator.JoyYRaw_ANA2, RawButton := bench.Operator.JoyBtnRaw, Cfg := cfg, NeutralXMem := nx, NeutralYMem := ny);
home(DeadmanArmed := joy.DeadmanArmed, JoystickDeflected := NOT joy.AtNeutralXY, JoystickPull := joy.AxisCmdY.DirectionPositive, JoystickPush := joy.AxisCmdY.DirectionNegative, BtnValidation := bench.Operator.JoyBtnRaw);
IF bench.Operator.JoyBtnRaw AND NOT previousButton THEN buttonEdges := buttonEdges + 1; END_IF; previousButton := bench.Operator.JoyBtnRaw;
ASSERT_FALSE(joy.DeadmanArmed, 'Maintien reel superieur a appui simule donc refus'); ASSERT_FALSE(joy.AxisCmdX.StartStop, 'Aucun bypass');
ADVANCE_TIME(10000000);
bench(RawPosM1 := raw1, RawPosM2 := raw2);
joy(RawX := bench.Operator.JoyXRaw_ANA1, RawY := bench.Operator.JoyYRaw_ANA2, RawButton := bench.Operator.JoyBtnRaw, Cfg := cfg, NeutralXMem := nx, NeutralYMem := ny);
home(DeadmanArmed := joy.DeadmanArmed, JoystickDeflected := NOT joy.AtNeutralXY, JoystickPull := joy.AxisCmdY.DirectionPositive, JoystickPush := joy.AxisCmdY.DirectionNegative, BtnValidation := bench.Operator.JoyBtnRaw);
IF bench.Operator.JoyBtnRaw AND NOT previousButton THEN buttonEdges := buttonEdges + 1; END_IF; previousButton := bench.Operator.JoyBtnRaw;
ASSERT_FALSE(joy.DeadmanArmed, 'Maintien reel superieur a appui simule donc refus'); ASSERT_FALSE(joy.AxisCmdX.StartStop, 'Aucun bypass');
ADVANCE_TIME(10000000);
bench(RawPosM1 := raw1, RawPosM2 := raw2);
joy(RawX := bench.Operator.JoyXRaw_ANA1, RawY := bench.Operator.JoyYRaw_ANA2, RawButton := bench.Operator.JoyBtnRaw, Cfg := cfg, NeutralXMem := nx, NeutralYMem := ny);
home(DeadmanArmed := joy.DeadmanArmed, JoystickDeflected := NOT joy.AtNeutralXY, JoystickPull := joy.AxisCmdY.DirectionPositive, JoystickPush := joy.AxisCmdY.DirectionNegative, BtnValidation := bench.Operator.JoyBtnRaw);
IF bench.Operator.JoyBtnRaw AND NOT previousButton THEN buttonEdges := buttonEdges + 1; END_IF; previousButton := bench.Operator.JoyBtnRaw;
ASSERT_FALSE(joy.DeadmanArmed, 'Maintien reel superieur a appui simule donc refus'); ASSERT_FALSE(joy.AxisCmdX.StartStop, 'Aucun bypass');
ADVANCE_TIME(10000000);
bench(RawPosM1 := raw1, RawPosM2 := raw2);
joy(RawX := bench.Operator.JoyXRaw_ANA1, RawY := bench.Operator.JoyYRaw_ANA2, RawButton := bench.Operator.JoyBtnRaw, Cfg := cfg, NeutralXMem := nx, NeutralYMem := ny);
home(DeadmanArmed := joy.DeadmanArmed, JoystickDeflected := NOT joy.AtNeutralXY, JoystickPull := joy.AxisCmdY.DirectionPositive, JoystickPush := joy.AxisCmdY.DirectionNegative, BtnValidation := bench.Operator.JoyBtnRaw);
IF bench.Operator.JoyBtnRaw AND NOT previousButton THEN buttonEdges := buttonEdges + 1; END_IF; previousButton := bench.Operator.JoyBtnRaw;
ASSERT_FALSE(joy.DeadmanArmed, 'Maintien reel superieur a appui simule donc refus'); ASSERT_FALSE(joy.AxisCmdX.StartStop, 'Aucun bypass');
ADVANCE_TIME(10000000);
bench(RawPosM1 := raw1, RawPosM2 := raw2);
joy(RawX := bench.Operator.JoyXRaw_ANA1, RawY := bench.Operator.JoyYRaw_ANA2, RawButton := bench.Operator.JoyBtnRaw, Cfg := cfg, NeutralXMem := nx, NeutralYMem := ny);
home(DeadmanArmed := joy.DeadmanArmed, JoystickDeflected := NOT joy.AtNeutralXY, JoystickPull := joy.AxisCmdY.DirectionPositive, JoystickPush := joy.AxisCmdY.DirectionNegative, BtnValidation := bench.Operator.JoyBtnRaw);
IF bench.Operator.JoyBtnRaw AND NOT previousButton THEN buttonEdges := buttonEdges + 1; END_IF; previousButton := bench.Operator.JoyBtnRaw;
ASSERT_FALSE(joy.DeadmanArmed, 'Maintien reel superieur a appui simule donc refus'); ASSERT_FALSE(joy.AxisCmdX.StartStop, 'Aucun bypass');
END_TEST

TEST 'TC-T418-INT-008 Bascule source reinitialise geste et refuse reprise tenue'
nx := 5000; ny := 5000; raw1 := 0; raw2 := 0; previousButton := FALSE; buttonEdges := 0;
bench.Enable := TRUE; joy.Enable := TRUE; joy.ArmingPermit := TRUE; diagOk.Operational := TRUE; joy.BusCanOpenOP := diagOk; joy.JoystickOP := diagOk; sourceSelected := TRUE; bench.HwReal.Operator.JoyXRaw_ANA1 := 5000; bench.HwReal.Operator.JoyYRaw_ANA2 := 5000;
ADVANCE_TIME(10000000); bench.OperatorSourceActive := sourceSelected; bench(RawPosM1 := raw1, RawPosM2 := raw2);
IF sourceSelected THEN selectedX := bench.Operator.JoyXRaw_ANA1; selectedY := bench.Operator.JoyYRaw_ANA2; selectedButton := bench.Operator.JoyBtnRaw; ELSE selectedX := 5000; selectedY := 5000; selectedButton := FALSE; END_IF;
joy(RawX := selectedX, RawY := selectedY, RawButton := selectedButton, Cfg := cfg, NeutralXMem := nx, NeutralYMem := ny);
IF bench.Operator.JoyBtnRaw AND NOT previousButton THEN buttonEdges := buttonEdges + 1; END_IF; previousButton := bench.Operator.JoyBtnRaw;
bench.SimJoystickRight_Fwd_MAINT_Active := TRUE;
ADVANCE_TIME(10000000); bench.OperatorSourceActive := sourceSelected; bench(RawPosM1 := raw1, RawPosM2 := raw2);
IF sourceSelected THEN selectedX := bench.Operator.JoyXRaw_ANA1; selectedY := bench.Operator.JoyYRaw_ANA2; selectedButton := bench.Operator.JoyBtnRaw; ELSE selectedX := 5000; selectedY := 5000; selectedButton := FALSE; END_IF;
joy(RawX := selectedX, RawY := selectedY, RawButton := selectedButton, Cfg := cfg, NeutralXMem := nx, NeutralYMem := ny);
IF bench.Operator.JoyBtnRaw AND NOT previousButton THEN buttonEdges := buttonEdges + 1; END_IF; previousButton := bench.Operator.JoyBtnRaw;
ADVANCE_TIME(10000000); bench.OperatorSourceActive := sourceSelected; bench(RawPosM1 := raw1, RawPosM2 := raw2);
IF sourceSelected THEN selectedX := bench.Operator.JoyXRaw_ANA1; selectedY := bench.Operator.JoyYRaw_ANA2; selectedButton := bench.Operator.JoyBtnRaw; ELSE selectedX := 5000; selectedY := 5000; selectedButton := FALSE; END_IF;
joy(RawX := selectedX, RawY := selectedY, RawButton := selectedButton, Cfg := cfg, NeutralXMem := nx, NeutralYMem := ny);
IF bench.Operator.JoyBtnRaw AND NOT previousButton THEN buttonEdges := buttonEdges + 1; END_IF; previousButton := bench.Operator.JoyBtnRaw;
ADVANCE_TIME(10000000); bench.OperatorSourceActive := sourceSelected; bench(RawPosM1 := raw1, RawPosM2 := raw2);
IF sourceSelected THEN selectedX := bench.Operator.JoyXRaw_ANA1; selectedY := bench.Operator.JoyYRaw_ANA2; selectedButton := bench.Operator.JoyBtnRaw; ELSE selectedX := 5000; selectedY := 5000; selectedButton := FALSE; END_IF;
joy(RawX := selectedX, RawY := selectedY, RawButton := selectedButton, Cfg := cfg, NeutralXMem := nx, NeutralYMem := ny);
IF bench.Operator.JoyBtnRaw AND NOT previousButton THEN buttonEdges := buttonEdges + 1; END_IF; previousButton := bench.Operator.JoyBtnRaw;
ADVANCE_TIME(10000000); bench.OperatorSourceActive := sourceSelected; bench(RawPosM1 := raw1, RawPosM2 := raw2);
IF sourceSelected THEN selectedX := bench.Operator.JoyXRaw_ANA1; selectedY := bench.Operator.JoyYRaw_ANA2; selectedButton := bench.Operator.JoyBtnRaw; ELSE selectedX := 5000; selectedY := 5000; selectedButton := FALSE; END_IF;
joy(RawX := selectedX, RawY := selectedY, RawButton := selectedButton, Cfg := cfg, NeutralXMem := nx, NeutralYMem := ny);
IF bench.Operator.JoyBtnRaw AND NOT previousButton THEN buttonEdges := buttonEdges + 1; END_IF; previousButton := bench.Operator.JoyBtnRaw;
ADVANCE_TIME(10000000); bench.OperatorSourceActive := sourceSelected; bench(RawPosM1 := raw1, RawPosM2 := raw2);
IF sourceSelected THEN selectedX := bench.Operator.JoyXRaw_ANA1; selectedY := bench.Operator.JoyYRaw_ANA2; selectedButton := bench.Operator.JoyBtnRaw; ELSE selectedX := 5000; selectedY := 5000; selectedButton := FALSE; END_IF;
joy(RawX := selectedX, RawY := selectedY, RawButton := selectedButton, Cfg := cfg, NeutralXMem := nx, NeutralYMem := ny);
IF bench.Operator.JoyBtnRaw AND NOT previousButton THEN buttonEdges := buttonEdges + 1; END_IF; previousButton := bench.Operator.JoyBtnRaw;
ADVANCE_TIME(10000000); bench.OperatorSourceActive := sourceSelected; bench(RawPosM1 := raw1, RawPosM2 := raw2);
IF sourceSelected THEN selectedX := bench.Operator.JoyXRaw_ANA1; selectedY := bench.Operator.JoyYRaw_ANA2; selectedButton := bench.Operator.JoyBtnRaw; ELSE selectedX := 5000; selectedY := 5000; selectedButton := FALSE; END_IF;
joy(RawX := selectedX, RawY := selectedY, RawButton := selectedButton, Cfg := cfg, NeutralXMem := nx, NeutralYMem := ny);
IF bench.Operator.JoyBtnRaw AND NOT previousButton THEN buttonEdges := buttonEdges + 1; END_IF; previousButton := bench.Operator.JoyBtnRaw;
ADVANCE_TIME(10000000); bench.OperatorSourceActive := sourceSelected; bench(RawPosM1 := raw1, RawPosM2 := raw2);
IF sourceSelected THEN selectedX := bench.Operator.JoyXRaw_ANA1; selectedY := bench.Operator.JoyYRaw_ANA2; selectedButton := bench.Operator.JoyBtnRaw; ELSE selectedX := 5000; selectedY := 5000; selectedButton := FALSE; END_IF;
joy(RawX := selectedX, RawY := selectedY, RawButton := selectedButton, Cfg := cfg, NeutralXMem := nx, NeutralYMem := ny);
IF bench.Operator.JoyBtnRaw AND NOT previousButton THEN buttonEdges := buttonEdges + 1; END_IF; previousButton := bench.Operator.JoyBtnRaw;
ADVANCE_TIME(10000000); bench.OperatorSourceActive := sourceSelected; bench(RawPosM1 := raw1, RawPosM2 := raw2);
IF sourceSelected THEN selectedX := bench.Operator.JoyXRaw_ANA1; selectedY := bench.Operator.JoyYRaw_ANA2; selectedButton := bench.Operator.JoyBtnRaw; ELSE selectedX := 5000; selectedY := 5000; selectedButton := FALSE; END_IF;
joy(RawX := selectedX, RawY := selectedY, RawButton := selectedButton, Cfg := cfg, NeutralXMem := nx, NeutralYMem := ny);
IF bench.Operator.JoyBtnRaw AND NOT previousButton THEN buttonEdges := buttonEdges + 1; END_IF; previousButton := bench.Operator.JoyBtnRaw;
ADVANCE_TIME(10000000); bench.OperatorSourceActive := sourceSelected; bench(RawPosM1 := raw1, RawPosM2 := raw2);
IF sourceSelected THEN selectedX := bench.Operator.JoyXRaw_ANA1; selectedY := bench.Operator.JoyYRaw_ANA2; selectedButton := bench.Operator.JoyBtnRaw; ELSE selectedX := 5000; selectedY := 5000; selectedButton := FALSE; END_IF;
joy(RawX := selectedX, RawY := selectedY, RawButton := selectedButton, Cfg := cfg, NeutralXMem := nx, NeutralYMem := ny);
IF bench.Operator.JoyBtnRaw AND NOT previousButton THEN buttonEdges := buttonEdges + 1; END_IF; previousButton := bench.Operator.JoyBtnRaw;
ADVANCE_TIME(10000000); bench.OperatorSourceActive := sourceSelected; bench(RawPosM1 := raw1, RawPosM2 := raw2);
IF sourceSelected THEN selectedX := bench.Operator.JoyXRaw_ANA1; selectedY := bench.Operator.JoyYRaw_ANA2; selectedButton := bench.Operator.JoyBtnRaw; ELSE selectedX := 5000; selectedY := 5000; selectedButton := FALSE; END_IF;
joy(RawX := selectedX, RawY := selectedY, RawButton := selectedButton, Cfg := cfg, NeutralXMem := nx, NeutralYMem := ny);
IF bench.Operator.JoyBtnRaw AND NOT previousButton THEN buttonEdges := buttonEdges + 1; END_IF; previousButton := bench.Operator.JoyBtnRaw;
ADVANCE_TIME(10000000); bench.OperatorSourceActive := sourceSelected; bench(RawPosM1 := raw1, RawPosM2 := raw2);
IF sourceSelected THEN selectedX := bench.Operator.JoyXRaw_ANA1; selectedY := bench.Operator.JoyYRaw_ANA2; selectedButton := bench.Operator.JoyBtnRaw; ELSE selectedX := 5000; selectedY := 5000; selectedButton := FALSE; END_IF;
joy(RawX := selectedX, RawY := selectedY, RawButton := selectedButton, Cfg := cfg, NeutralXMem := nx, NeutralYMem := ny);
IF bench.Operator.JoyBtnRaw AND NOT previousButton THEN buttonEdges := buttonEdges + 1; END_IF; previousButton := bench.Operator.JoyBtnRaw;
ADVANCE_TIME(10000000); bench.OperatorSourceActive := sourceSelected; bench(RawPosM1 := raw1, RawPosM2 := raw2);
IF sourceSelected THEN selectedX := bench.Operator.JoyXRaw_ANA1; selectedY := bench.Operator.JoyYRaw_ANA2; selectedButton := bench.Operator.JoyBtnRaw; ELSE selectedX := 5000; selectedY := 5000; selectedButton := FALSE; END_IF;
joy(RawX := selectedX, RawY := selectedY, RawButton := selectedButton, Cfg := cfg, NeutralXMem := nx, NeutralYMem := ny);
IF bench.Operator.JoyBtnRaw AND NOT previousButton THEN buttonEdges := buttonEdges + 1; END_IF; previousButton := bench.Operator.JoyBtnRaw;
ADVANCE_TIME(10000000); bench.OperatorSourceActive := sourceSelected; bench(RawPosM1 := raw1, RawPosM2 := raw2);
IF sourceSelected THEN selectedX := bench.Operator.JoyXRaw_ANA1; selectedY := bench.Operator.JoyYRaw_ANA2; selectedButton := bench.Operator.JoyBtnRaw; ELSE selectedX := 5000; selectedY := 5000; selectedButton := FALSE; END_IF;
joy(RawX := selectedX, RawY := selectedY, RawButton := selectedButton, Cfg := cfg, NeutralXMem := nx, NeutralYMem := ny);
IF bench.Operator.JoyBtnRaw AND NOT previousButton THEN buttonEdges := buttonEdges + 1; END_IF; previousButton := bench.Operator.JoyBtnRaw;
ADVANCE_TIME(10000000); bench.OperatorSourceActive := sourceSelected; bench(RawPosM1 := raw1, RawPosM2 := raw2);
IF sourceSelected THEN selectedX := bench.Operator.JoyXRaw_ANA1; selectedY := bench.Operator.JoyYRaw_ANA2; selectedButton := bench.Operator.JoyBtnRaw; ELSE selectedX := 5000; selectedY := 5000; selectedButton := FALSE; END_IF;
joy(RawX := selectedX, RawY := selectedY, RawButton := selectedButton, Cfg := cfg, NeutralXMem := nx, NeutralYMem := ny);
IF bench.Operator.JoyBtnRaw AND NOT previousButton THEN buttonEdges := buttonEdges + 1; END_IF; previousButton := bench.Operator.JoyBtnRaw;
ADVANCE_TIME(10000000); bench.OperatorSourceActive := sourceSelected; bench(RawPosM1 := raw1, RawPosM2 := raw2);
IF sourceSelected THEN selectedX := bench.Operator.JoyXRaw_ANA1; selectedY := bench.Operator.JoyYRaw_ANA2; selectedButton := bench.Operator.JoyBtnRaw; ELSE selectedX := 5000; selectedY := 5000; selectedButton := FALSE; END_IF;
joy(RawX := selectedX, RawY := selectedY, RawButton := selectedButton, Cfg := cfg, NeutralXMem := nx, NeutralYMem := ny);
IF bench.Operator.JoyBtnRaw AND NOT previousButton THEN buttonEdges := buttonEdges + 1; END_IF; previousButton := bench.Operator.JoyBtnRaw;
ADVANCE_TIME(10000000); bench.OperatorSourceActive := sourceSelected; bench(RawPosM1 := raw1, RawPosM2 := raw2);
IF sourceSelected THEN selectedX := bench.Operator.JoyXRaw_ANA1; selectedY := bench.Operator.JoyYRaw_ANA2; selectedButton := bench.Operator.JoyBtnRaw; ELSE selectedX := 5000; selectedY := 5000; selectedButton := FALSE; END_IF;
joy(RawX := selectedX, RawY := selectedY, RawButton := selectedButton, Cfg := cfg, NeutralXMem := nx, NeutralYMem := ny);
IF bench.Operator.JoyBtnRaw AND NOT previousButton THEN buttonEdges := buttonEdges + 1; END_IF; previousButton := bench.Operator.JoyBtnRaw;
ADVANCE_TIME(10000000); bench.OperatorSourceActive := sourceSelected; bench(RawPosM1 := raw1, RawPosM2 := raw2);
IF sourceSelected THEN selectedX := bench.Operator.JoyXRaw_ANA1; selectedY := bench.Operator.JoyYRaw_ANA2; selectedButton := bench.Operator.JoyBtnRaw; ELSE selectedX := 5000; selectedY := 5000; selectedButton := FALSE; END_IF;
joy(RawX := selectedX, RawY := selectedY, RawButton := selectedButton, Cfg := cfg, NeutralXMem := nx, NeutralYMem := ny);
IF bench.Operator.JoyBtnRaw AND NOT previousButton THEN buttonEdges := buttonEdges + 1; END_IF; previousButton := bench.Operator.JoyBtnRaw;
ADVANCE_TIME(10000000); bench.OperatorSourceActive := sourceSelected; bench(RawPosM1 := raw1, RawPosM2 := raw2);
IF sourceSelected THEN selectedX := bench.Operator.JoyXRaw_ANA1; selectedY := bench.Operator.JoyYRaw_ANA2; selectedButton := bench.Operator.JoyBtnRaw; ELSE selectedX := 5000; selectedY := 5000; selectedButton := FALSE; END_IF;
joy(RawX := selectedX, RawY := selectedY, RawButton := selectedButton, Cfg := cfg, NeutralXMem := nx, NeutralYMem := ny);
IF bench.Operator.JoyBtnRaw AND NOT previousButton THEN buttonEdges := buttonEdges + 1; END_IF; previousButton := bench.Operator.JoyBtnRaw;
ADVANCE_TIME(10000000); bench.OperatorSourceActive := sourceSelected; bench(RawPosM1 := raw1, RawPosM2 := raw2);
IF sourceSelected THEN selectedX := bench.Operator.JoyXRaw_ANA1; selectedY := bench.Operator.JoyYRaw_ANA2; selectedButton := bench.Operator.JoyBtnRaw; ELSE selectedX := 5000; selectedY := 5000; selectedButton := FALSE; END_IF;
joy(RawX := selectedX, RawY := selectedY, RawButton := selectedButton, Cfg := cfg, NeutralXMem := nx, NeutralYMem := ny);
IF bench.Operator.JoyBtnRaw AND NOT previousButton THEN buttonEdges := buttonEdges + 1; END_IF; previousButton := bench.Operator.JoyBtnRaw;
ADVANCE_TIME(10000000); bench.OperatorSourceActive := sourceSelected; bench(RawPosM1 := raw1, RawPosM2 := raw2);
IF sourceSelected THEN selectedX := bench.Operator.JoyXRaw_ANA1; selectedY := bench.Operator.JoyYRaw_ANA2; selectedButton := bench.Operator.JoyBtnRaw; ELSE selectedX := 5000; selectedY := 5000; selectedButton := FALSE; END_IF;
joy(RawX := selectedX, RawY := selectedY, RawButton := selectedButton, Cfg := cfg, NeutralXMem := nx, NeutralYMem := ny);
IF bench.Operator.JoyBtnRaw AND NOT previousButton THEN buttonEdges := buttonEdges + 1; END_IF; previousButton := bench.Operator.JoyBtnRaw;
ADVANCE_TIME(10000000); bench.OperatorSourceActive := sourceSelected; bench(RawPosM1 := raw1, RawPosM2 := raw2);
IF sourceSelected THEN selectedX := bench.Operator.JoyXRaw_ANA1; selectedY := bench.Operator.JoyYRaw_ANA2; selectedButton := bench.Operator.JoyBtnRaw; ELSE selectedX := 5000; selectedY := 5000; selectedButton := FALSE; END_IF;
joy(RawX := selectedX, RawY := selectedY, RawButton := selectedButton, Cfg := cfg, NeutralXMem := nx, NeutralYMem := ny);
IF bench.Operator.JoyBtnRaw AND NOT previousButton THEN buttonEdges := buttonEdges + 1; END_IF; previousButton := bench.Operator.JoyBtnRaw;
ADVANCE_TIME(10000000); bench.OperatorSourceActive := sourceSelected; bench(RawPosM1 := raw1, RawPosM2 := raw2);
IF sourceSelected THEN selectedX := bench.Operator.JoyXRaw_ANA1; selectedY := bench.Operator.JoyYRaw_ANA2; selectedButton := bench.Operator.JoyBtnRaw; ELSE selectedX := 5000; selectedY := 5000; selectedButton := FALSE; END_IF;
joy(RawX := selectedX, RawY := selectedY, RawButton := selectedButton, Cfg := cfg, NeutralXMem := nx, NeutralYMem := ny);
IF bench.Operator.JoyBtnRaw AND NOT previousButton THEN buttonEdges := buttonEdges + 1; END_IF; previousButton := bench.Operator.JoyBtnRaw;
ADVANCE_TIME(10000000); bench.OperatorSourceActive := sourceSelected; bench(RawPosM1 := raw1, RawPosM2 := raw2);
IF sourceSelected THEN selectedX := bench.Operator.JoyXRaw_ANA1; selectedY := bench.Operator.JoyYRaw_ANA2; selectedButton := bench.Operator.JoyBtnRaw; ELSE selectedX := 5000; selectedY := 5000; selectedButton := FALSE; END_IF;
joy(RawX := selectedX, RawY := selectedY, RawButton := selectedButton, Cfg := cfg, NeutralXMem := nx, NeutralYMem := ny);
IF bench.Operator.JoyBtnRaw AND NOT previousButton THEN buttonEdges := buttonEdges + 1; END_IF; previousButton := bench.Operator.JoyBtnRaw;
ADVANCE_TIME(10000000); bench.OperatorSourceActive := sourceSelected; bench(RawPosM1 := raw1, RawPosM2 := raw2);
IF sourceSelected THEN selectedX := bench.Operator.JoyXRaw_ANA1; selectedY := bench.Operator.JoyYRaw_ANA2; selectedButton := bench.Operator.JoyBtnRaw; ELSE selectedX := 5000; selectedY := 5000; selectedButton := FALSE; END_IF;
joy(RawX := selectedX, RawY := selectedY, RawButton := selectedButton, Cfg := cfg, NeutralXMem := nx, NeutralYMem := ny);
IF bench.Operator.JoyBtnRaw AND NOT previousButton THEN buttonEdges := buttonEdges + 1; END_IF; previousButton := bench.Operator.JoyBtnRaw;
ADVANCE_TIME(10000000); bench.OperatorSourceActive := sourceSelected; bench(RawPosM1 := raw1, RawPosM2 := raw2);
IF sourceSelected THEN selectedX := bench.Operator.JoyXRaw_ANA1; selectedY := bench.Operator.JoyYRaw_ANA2; selectedButton := bench.Operator.JoyBtnRaw; ELSE selectedX := 5000; selectedY := 5000; selectedButton := FALSE; END_IF;
joy(RawX := selectedX, RawY := selectedY, RawButton := selectedButton, Cfg := cfg, NeutralXMem := nx, NeutralYMem := ny);
IF bench.Operator.JoyBtnRaw AND NOT previousButton THEN buttonEdges := buttonEdges + 1; END_IF; previousButton := bench.Operator.JoyBtnRaw;
ADVANCE_TIME(10000000); bench.OperatorSourceActive := sourceSelected; bench(RawPosM1 := raw1, RawPosM2 := raw2);
IF sourceSelected THEN selectedX := bench.Operator.JoyXRaw_ANA1; selectedY := bench.Operator.JoyYRaw_ANA2; selectedButton := bench.Operator.JoyBtnRaw; ELSE selectedX := 5000; selectedY := 5000; selectedButton := FALSE; END_IF;
joy(RawX := selectedX, RawY := selectedY, RawButton := selectedButton, Cfg := cfg, NeutralXMem := nx, NeutralYMem := ny);
IF bench.Operator.JoyBtnRaw AND NOT previousButton THEN buttonEdges := buttonEdges + 1; END_IF; previousButton := bench.Operator.JoyBtnRaw;
ADVANCE_TIME(10000000); bench.OperatorSourceActive := sourceSelected; bench(RawPosM1 := raw1, RawPosM2 := raw2);
IF sourceSelected THEN selectedX := bench.Operator.JoyXRaw_ANA1; selectedY := bench.Operator.JoyYRaw_ANA2; selectedButton := bench.Operator.JoyBtnRaw; ELSE selectedX := 5000; selectedY := 5000; selectedButton := FALSE; END_IF;
joy(RawX := selectedX, RawY := selectedY, RawButton := selectedButton, Cfg := cfg, NeutralXMem := nx, NeutralYMem := ny);
IF bench.Operator.JoyBtnRaw AND NOT previousButton THEN buttonEdges := buttonEdges + 1; END_IF; previousButton := bench.Operator.JoyBtnRaw;
ADVANCE_TIME(10000000); bench.OperatorSourceActive := sourceSelected; bench(RawPosM1 := raw1, RawPosM2 := raw2);
IF sourceSelected THEN selectedX := bench.Operator.JoyXRaw_ANA1; selectedY := bench.Operator.JoyYRaw_ANA2; selectedButton := bench.Operator.JoyBtnRaw; ELSE selectedX := 5000; selectedY := 5000; selectedButton := FALSE; END_IF;
joy(RawX := selectedX, RawY := selectedY, RawButton := selectedButton, Cfg := cfg, NeutralXMem := nx, NeutralYMem := ny);
IF bench.Operator.JoyBtnRaw AND NOT previousButton THEN buttonEdges := buttonEdges + 1; END_IF; previousButton := bench.Operator.JoyBtnRaw;
ADVANCE_TIME(10000000); bench.OperatorSourceActive := sourceSelected; bench(RawPosM1 := raw1, RawPosM2 := raw2);
IF sourceSelected THEN selectedX := bench.Operator.JoyXRaw_ANA1; selectedY := bench.Operator.JoyYRaw_ANA2; selectedButton := bench.Operator.JoyBtnRaw; ELSE selectedX := 5000; selectedY := 5000; selectedButton := FALSE; END_IF;
joy(RawX := selectedX, RawY := selectedY, RawButton := selectedButton, Cfg := cfg, NeutralXMem := nx, NeutralYMem := ny);
IF bench.Operator.JoyBtnRaw AND NOT previousButton THEN buttonEdges := buttonEdges + 1; END_IF; previousButton := bench.Operator.JoyBtnRaw;
ADVANCE_TIME(10000000); bench.OperatorSourceActive := sourceSelected; bench(RawPosM1 := raw1, RawPosM2 := raw2);
IF sourceSelected THEN selectedX := bench.Operator.JoyXRaw_ANA1; selectedY := bench.Operator.JoyYRaw_ANA2; selectedButton := bench.Operator.JoyBtnRaw; ELSE selectedX := 5000; selectedY := 5000; selectedButton := FALSE; END_IF;
joy(RawX := selectedX, RawY := selectedY, RawButton := selectedButton, Cfg := cfg, NeutralXMem := nx, NeutralYMem := ny);
IF bench.Operator.JoyBtnRaw AND NOT previousButton THEN buttonEdges := buttonEdges + 1; END_IF; previousButton := bench.Operator.JoyBtnRaw;
ADVANCE_TIME(10000000); bench.OperatorSourceActive := sourceSelected; bench(RawPosM1 := raw1, RawPosM2 := raw2);
IF sourceSelected THEN selectedX := bench.Operator.JoyXRaw_ANA1; selectedY := bench.Operator.JoyYRaw_ANA2; selectedButton := bench.Operator.JoyBtnRaw; ELSE selectedX := 5000; selectedY := 5000; selectedButton := FALSE; END_IF;
joy(RawX := selectedX, RawY := selectedY, RawButton := selectedButton, Cfg := cfg, NeutralXMem := nx, NeutralYMem := ny);
IF bench.Operator.JoyBtnRaw AND NOT previousButton THEN buttonEdges := buttonEdges + 1; END_IF; previousButton := bench.Operator.JoyBtnRaw;
ADVANCE_TIME(10000000); bench.OperatorSourceActive := sourceSelected; bench(RawPosM1 := raw1, RawPosM2 := raw2);
IF sourceSelected THEN selectedX := bench.Operator.JoyXRaw_ANA1; selectedY := bench.Operator.JoyYRaw_ANA2; selectedButton := bench.Operator.JoyBtnRaw; ELSE selectedX := 5000; selectedY := 5000; selectedButton := FALSE; END_IF;
joy(RawX := selectedX, RawY := selectedY, RawButton := selectedButton, Cfg := cfg, NeutralXMem := nx, NeutralYMem := ny);
IF bench.Operator.JoyBtnRaw AND NOT previousButton THEN buttonEdges := buttonEdges + 1; END_IF; previousButton := bench.Operator.JoyBtnRaw;
ADVANCE_TIME(10000000); bench.OperatorSourceActive := sourceSelected; bench(RawPosM1 := raw1, RawPosM2 := raw2);
IF sourceSelected THEN selectedX := bench.Operator.JoyXRaw_ANA1; selectedY := bench.Operator.JoyYRaw_ANA2; selectedButton := bench.Operator.JoyBtnRaw; ELSE selectedX := 5000; selectedY := 5000; selectedButton := FALSE; END_IF;
joy(RawX := selectedX, RawY := selectedY, RawButton := selectedButton, Cfg := cfg, NeutralXMem := nx, NeutralYMem := ny);
IF bench.Operator.JoyBtnRaw AND NOT previousButton THEN buttonEdges := buttonEdges + 1; END_IF; previousButton := bench.Operator.JoyBtnRaw;
ADVANCE_TIME(10000000); bench.OperatorSourceActive := sourceSelected; bench(RawPosM1 := raw1, RawPosM2 := raw2);
IF sourceSelected THEN selectedX := bench.Operator.JoyXRaw_ANA1; selectedY := bench.Operator.JoyYRaw_ANA2; selectedButton := bench.Operator.JoyBtnRaw; ELSE selectedX := 5000; selectedY := 5000; selectedButton := FALSE; END_IF;
joy(RawX := selectedX, RawY := selectedY, RawButton := selectedButton, Cfg := cfg, NeutralXMem := nx, NeutralYMem := ny);
IF bench.Operator.JoyBtnRaw AND NOT previousButton THEN buttonEdges := buttonEdges + 1; END_IF; previousButton := bench.Operator.JoyBtnRaw;
ADVANCE_TIME(10000000); bench.OperatorSourceActive := sourceSelected; bench(RawPosM1 := raw1, RawPosM2 := raw2);
IF sourceSelected THEN selectedX := bench.Operator.JoyXRaw_ANA1; selectedY := bench.Operator.JoyYRaw_ANA2; selectedButton := bench.Operator.JoyBtnRaw; ELSE selectedX := 5000; selectedY := 5000; selectedButton := FALSE; END_IF;
joy(RawX := selectedX, RawY := selectedY, RawButton := selectedButton, Cfg := cfg, NeutralXMem := nx, NeutralYMem := ny);
IF bench.Operator.JoyBtnRaw AND NOT previousButton THEN buttonEdges := buttonEdges + 1; END_IF; previousButton := bench.Operator.JoyBtnRaw;
ADVANCE_TIME(10000000); bench.OperatorSourceActive := sourceSelected; bench(RawPosM1 := raw1, RawPosM2 := raw2);
IF sourceSelected THEN selectedX := bench.Operator.JoyXRaw_ANA1; selectedY := bench.Operator.JoyYRaw_ANA2; selectedButton := bench.Operator.JoyBtnRaw; ELSE selectedX := 5000; selectedY := 5000; selectedButton := FALSE; END_IF;
joy(RawX := selectedX, RawY := selectedY, RawButton := selectedButton, Cfg := cfg, NeutralXMem := nx, NeutralYMem := ny);
IF bench.Operator.JoyBtnRaw AND NOT previousButton THEN buttonEdges := buttonEdges + 1; END_IF; previousButton := bench.Operator.JoyBtnRaw;
ADVANCE_TIME(10000000); bench.OperatorSourceActive := sourceSelected; bench(RawPosM1 := raw1, RawPosM2 := raw2);
IF sourceSelected THEN selectedX := bench.Operator.JoyXRaw_ANA1; selectedY := bench.Operator.JoyYRaw_ANA2; selectedButton := bench.Operator.JoyBtnRaw; ELSE selectedX := 5000; selectedY := 5000; selectedButton := FALSE; END_IF;
joy(RawX := selectedX, RawY := selectedY, RawButton := selectedButton, Cfg := cfg, NeutralXMem := nx, NeutralYMem := ny);
IF bench.Operator.JoyBtnRaw AND NOT previousButton THEN buttonEdges := buttonEdges + 1; END_IF; previousButton := bench.Operator.JoyBtnRaw;
ADVANCE_TIME(10000000); bench.OperatorSourceActive := sourceSelected; bench(RawPosM1 := raw1, RawPosM2 := raw2);
IF sourceSelected THEN selectedX := bench.Operator.JoyXRaw_ANA1; selectedY := bench.Operator.JoyYRaw_ANA2; selectedButton := bench.Operator.JoyBtnRaw; ELSE selectedX := 5000; selectedY := 5000; selectedButton := FALSE; END_IF;
joy(RawX := selectedX, RawY := selectedY, RawButton := selectedButton, Cfg := cfg, NeutralXMem := nx, NeutralYMem := ny);
IF bench.Operator.JoyBtnRaw AND NOT previousButton THEN buttonEdges := buttonEdges + 1; END_IF; previousButton := bench.Operator.JoyBtnRaw;
ADVANCE_TIME(10000000); bench.OperatorSourceActive := sourceSelected; bench(RawPosM1 := raw1, RawPosM2 := raw2);
IF sourceSelected THEN selectedX := bench.Operator.JoyXRaw_ANA1; selectedY := bench.Operator.JoyYRaw_ANA2; selectedButton := bench.Operator.JoyBtnRaw; ELSE selectedX := 5000; selectedY := 5000; selectedButton := FALSE; END_IF;
joy(RawX := selectedX, RawY := selectedY, RawButton := selectedButton, Cfg := cfg, NeutralXMem := nx, NeutralYMem := ny);
IF bench.Operator.JoyBtnRaw AND NOT previousButton THEN buttonEdges := buttonEdges + 1; END_IF; previousButton := bench.Operator.JoyBtnRaw;
ADVANCE_TIME(10000000); bench.OperatorSourceActive := sourceSelected; bench(RawPosM1 := raw1, RawPosM2 := raw2);
IF sourceSelected THEN selectedX := bench.Operator.JoyXRaw_ANA1; selectedY := bench.Operator.JoyYRaw_ANA2; selectedButton := bench.Operator.JoyBtnRaw; ELSE selectedX := 5000; selectedY := 5000; selectedButton := FALSE; END_IF;
joy(RawX := selectedX, RawY := selectedY, RawButton := selectedButton, Cfg := cfg, NeutralXMem := nx, NeutralYMem := ny);
IF bench.Operator.JoyBtnRaw AND NOT previousButton THEN buttonEdges := buttonEdges + 1; END_IF; previousButton := bench.Operator.JoyBtnRaw;
ADVANCE_TIME(10000000); bench.OperatorSourceActive := sourceSelected; bench(RawPosM1 := raw1, RawPosM2 := raw2);
IF sourceSelected THEN selectedX := bench.Operator.JoyXRaw_ANA1; selectedY := bench.Operator.JoyYRaw_ANA2; selectedButton := bench.Operator.JoyBtnRaw; ELSE selectedX := 5000; selectedY := 5000; selectedButton := FALSE; END_IF;
joy(RawX := selectedX, RawY := selectedY, RawButton := selectedButton, Cfg := cfg, NeutralXMem := nx, NeutralYMem := ny);
IF bench.Operator.JoyBtnRaw AND NOT previousButton THEN buttonEdges := buttonEdges + 1; END_IF; previousButton := bench.Operator.JoyBtnRaw;
ADVANCE_TIME(10000000); bench.OperatorSourceActive := sourceSelected; bench(RawPosM1 := raw1, RawPosM2 := raw2);
IF sourceSelected THEN selectedX := bench.Operator.JoyXRaw_ANA1; selectedY := bench.Operator.JoyYRaw_ANA2; selectedButton := bench.Operator.JoyBtnRaw; ELSE selectedX := 5000; selectedY := 5000; selectedButton := FALSE; END_IF;
joy(RawX := selectedX, RawY := selectedY, RawButton := selectedButton, Cfg := cfg, NeutralXMem := nx, NeutralYMem := ny);
IF bench.Operator.JoyBtnRaw AND NOT previousButton THEN buttonEdges := buttonEdges + 1; END_IF; previousButton := bench.Operator.JoyBtnRaw;
ADVANCE_TIME(10000000); bench.OperatorSourceActive := sourceSelected; bench(RawPosM1 := raw1, RawPosM2 := raw2);
IF sourceSelected THEN selectedX := bench.Operator.JoyXRaw_ANA1; selectedY := bench.Operator.JoyYRaw_ANA2; selectedButton := bench.Operator.JoyBtnRaw; ELSE selectedX := 5000; selectedY := 5000; selectedButton := FALSE; END_IF;
joy(RawX := selectedX, RawY := selectedY, RawButton := selectedButton, Cfg := cfg, NeutralXMem := nx, NeutralYMem := ny);
IF bench.Operator.JoyBtnRaw AND NOT previousButton THEN buttonEdges := buttonEdges + 1; END_IF; previousButton := bench.Operator.JoyBtnRaw;
ADVANCE_TIME(10000000); bench.OperatorSourceActive := sourceSelected; bench(RawPosM1 := raw1, RawPosM2 := raw2);
IF sourceSelected THEN selectedX := bench.Operator.JoyXRaw_ANA1; selectedY := bench.Operator.JoyYRaw_ANA2; selectedButton := bench.Operator.JoyBtnRaw; ELSE selectedX := 5000; selectedY := 5000; selectedButton := FALSE; END_IF;
joy(RawX := selectedX, RawY := selectedY, RawButton := selectedButton, Cfg := cfg, NeutralXMem := nx, NeutralYMem := ny);
IF bench.Operator.JoyBtnRaw AND NOT previousButton THEN buttonEdges := buttonEdges + 1; END_IF; previousButton := bench.Operator.JoyBtnRaw;
ADVANCE_TIME(10000000); bench.OperatorSourceActive := sourceSelected; bench(RawPosM1 := raw1, RawPosM2 := raw2);
IF sourceSelected THEN selectedX := bench.Operator.JoyXRaw_ANA1; selectedY := bench.Operator.JoyYRaw_ANA2; selectedButton := bench.Operator.JoyBtnRaw; ELSE selectedX := 5000; selectedY := 5000; selectedButton := FALSE; END_IF;
joy(RawX := selectedX, RawY := selectedY, RawButton := selectedButton, Cfg := cfg, NeutralXMem := nx, NeutralYMem := ny);
IF bench.Operator.JoyBtnRaw AND NOT previousButton THEN buttonEdges := buttonEdges + 1; END_IF; previousButton := bench.Operator.JoyBtnRaw;
ADVANCE_TIME(10000000); bench.OperatorSourceActive := sourceSelected; bench(RawPosM1 := raw1, RawPosM2 := raw2);
IF sourceSelected THEN selectedX := bench.Operator.JoyXRaw_ANA1; selectedY := bench.Operator.JoyYRaw_ANA2; selectedButton := bench.Operator.JoyBtnRaw; ELSE selectedX := 5000; selectedY := 5000; selectedButton := FALSE; END_IF;
joy(RawX := selectedX, RawY := selectedY, RawButton := selectedButton, Cfg := cfg, NeutralXMem := nx, NeutralYMem := ny);
IF bench.Operator.JoyBtnRaw AND NOT previousButton THEN buttonEdges := buttonEdges + 1; END_IF; previousButton := bench.Operator.JoyBtnRaw;
ADVANCE_TIME(10000000); bench.OperatorSourceActive := sourceSelected; bench(RawPosM1 := raw1, RawPosM2 := raw2);
IF sourceSelected THEN selectedX := bench.Operator.JoyXRaw_ANA1; selectedY := bench.Operator.JoyYRaw_ANA2; selectedButton := bench.Operator.JoyBtnRaw; ELSE selectedX := 5000; selectedY := 5000; selectedButton := FALSE; END_IF;
joy(RawX := selectedX, RawY := selectedY, RawButton := selectedButton, Cfg := cfg, NeutralXMem := nx, NeutralYMem := ny);
IF bench.Operator.JoyBtnRaw AND NOT previousButton THEN buttonEdges := buttonEdges + 1; END_IF; previousButton := bench.Operator.JoyBtnRaw;
ADVANCE_TIME(10000000); bench.OperatorSourceActive := sourceSelected; bench(RawPosM1 := raw1, RawPosM2 := raw2);
IF sourceSelected THEN selectedX := bench.Operator.JoyXRaw_ANA1; selectedY := bench.Operator.JoyYRaw_ANA2; selectedButton := bench.Operator.JoyBtnRaw; ELSE selectedX := 5000; selectedY := 5000; selectedButton := FALSE; END_IF;
joy(RawX := selectedX, RawY := selectedY, RawButton := selectedButton, Cfg := cfg, NeutralXMem := nx, NeutralYMem := ny);
IF bench.Operator.JoyBtnRaw AND NOT previousButton THEN buttonEdges := buttonEdges + 1; END_IF; previousButton := bench.Operator.JoyBtnRaw;
ADVANCE_TIME(10000000); bench.OperatorSourceActive := sourceSelected; bench(RawPosM1 := raw1, RawPosM2 := raw2);
IF sourceSelected THEN selectedX := bench.Operator.JoyXRaw_ANA1; selectedY := bench.Operator.JoyYRaw_ANA2; selectedButton := bench.Operator.JoyBtnRaw; ELSE selectedX := 5000; selectedY := 5000; selectedButton := FALSE; END_IF;
joy(RawX := selectedX, RawY := selectedY, RawButton := selectedButton, Cfg := cfg, NeutralXMem := nx, NeutralYMem := ny);
IF bench.Operator.JoyBtnRaw AND NOT previousButton THEN buttonEdges := buttonEdges + 1; END_IF; previousButton := bench.Operator.JoyBtnRaw;
ADVANCE_TIME(10000000); bench.OperatorSourceActive := sourceSelected; bench(RawPosM1 := raw1, RawPosM2 := raw2);
IF sourceSelected THEN selectedX := bench.Operator.JoyXRaw_ANA1; selectedY := bench.Operator.JoyYRaw_ANA2; selectedButton := bench.Operator.JoyBtnRaw; ELSE selectedX := 5000; selectedY := 5000; selectedButton := FALSE; END_IF;
joy(RawX := selectedX, RawY := selectedY, RawButton := selectedButton, Cfg := cfg, NeutralXMem := nx, NeutralYMem := ny);
IF bench.Operator.JoyBtnRaw AND NOT previousButton THEN buttonEdges := buttonEdges + 1; END_IF; previousButton := bench.Operator.JoyBtnRaw;
ADVANCE_TIME(10000000); bench.OperatorSourceActive := sourceSelected; bench(RawPosM1 := raw1, RawPosM2 := raw2);
IF sourceSelected THEN selectedX := bench.Operator.JoyXRaw_ANA1; selectedY := bench.Operator.JoyYRaw_ANA2; selectedButton := bench.Operator.JoyBtnRaw; ELSE selectedX := 5000; selectedY := 5000; selectedButton := FALSE; END_IF;
joy(RawX := selectedX, RawY := selectedY, RawButton := selectedButton, Cfg := cfg, NeutralXMem := nx, NeutralYMem := ny);
IF bench.Operator.JoyBtnRaw AND NOT previousButton THEN buttonEdges := buttonEdges + 1; END_IF; previousButton := bench.Operator.JoyBtnRaw;
ADVANCE_TIME(10000000); bench.OperatorSourceActive := sourceSelected; bench(RawPosM1 := raw1, RawPosM2 := raw2);
IF sourceSelected THEN selectedX := bench.Operator.JoyXRaw_ANA1; selectedY := bench.Operator.JoyYRaw_ANA2; selectedButton := bench.Operator.JoyBtnRaw; ELSE selectedX := 5000; selectedY := 5000; selectedButton := FALSE; END_IF;
joy(RawX := selectedX, RawY := selectedY, RawButton := selectedButton, Cfg := cfg, NeutralXMem := nx, NeutralYMem := ny);
IF bench.Operator.JoyBtnRaw AND NOT previousButton THEN buttonEdges := buttonEdges + 1; END_IF; previousButton := bench.Operator.JoyBtnRaw;
ADVANCE_TIME(10000000); bench.OperatorSourceActive := sourceSelected; bench(RawPosM1 := raw1, RawPosM2 := raw2);
IF sourceSelected THEN selectedX := bench.Operator.JoyXRaw_ANA1; selectedY := bench.Operator.JoyYRaw_ANA2; selectedButton := bench.Operator.JoyBtnRaw; ELSE selectedX := 5000; selectedY := 5000; selectedButton := FALSE; END_IF;
joy(RawX := selectedX, RawY := selectedY, RawButton := selectedButton, Cfg := cfg, NeutralXMem := nx, NeutralYMem := ny);
IF bench.Operator.JoyBtnRaw AND NOT previousButton THEN buttonEdges := buttonEdges + 1; END_IF; previousButton := bench.Operator.JoyBtnRaw;
ADVANCE_TIME(10000000); bench.OperatorSourceActive := sourceSelected; bench(RawPosM1 := raw1, RawPosM2 := raw2);
IF sourceSelected THEN selectedX := bench.Operator.JoyXRaw_ANA1; selectedY := bench.Operator.JoyYRaw_ANA2; selectedButton := bench.Operator.JoyBtnRaw; ELSE selectedX := 5000; selectedY := 5000; selectedButton := FALSE; END_IF;
joy(RawX := selectedX, RawY := selectedY, RawButton := selectedButton, Cfg := cfg, NeutralXMem := nx, NeutralYMem := ny);
IF bench.Operator.JoyBtnRaw AND NOT previousButton THEN buttonEdges := buttonEdges + 1; END_IF; previousButton := bench.Operator.JoyBtnRaw;
ADVANCE_TIME(10000000); bench.OperatorSourceActive := sourceSelected; bench(RawPosM1 := raw1, RawPosM2 := raw2);
IF sourceSelected THEN selectedX := bench.Operator.JoyXRaw_ANA1; selectedY := bench.Operator.JoyYRaw_ANA2; selectedButton := bench.Operator.JoyBtnRaw; ELSE selectedX := 5000; selectedY := 5000; selectedButton := FALSE; END_IF;
joy(RawX := selectedX, RawY := selectedY, RawButton := selectedButton, Cfg := cfg, NeutralXMem := nx, NeutralYMem := ny);
IF bench.Operator.JoyBtnRaw AND NOT previousButton THEN buttonEdges := buttonEdges + 1; END_IF; previousButton := bench.Operator.JoyBtnRaw;
ADVANCE_TIME(10000000); bench.OperatorSourceActive := sourceSelected; bench(RawPosM1 := raw1, RawPosM2 := raw2);
IF sourceSelected THEN selectedX := bench.Operator.JoyXRaw_ANA1; selectedY := bench.Operator.JoyYRaw_ANA2; selectedButton := bench.Operator.JoyBtnRaw; ELSE selectedX := 5000; selectedY := 5000; selectedButton := FALSE; END_IF;
joy(RawX := selectedX, RawY := selectedY, RawButton := selectedButton, Cfg := cfg, NeutralXMem := nx, NeutralYMem := ny);
IF bench.Operator.JoyBtnRaw AND NOT previousButton THEN buttonEdges := buttonEdges + 1; END_IF; previousButton := bench.Operator.JoyBtnRaw;
ADVANCE_TIME(10000000); bench.OperatorSourceActive := sourceSelected; bench(RawPosM1 := raw1, RawPosM2 := raw2);
IF sourceSelected THEN selectedX := bench.Operator.JoyXRaw_ANA1; selectedY := bench.Operator.JoyYRaw_ANA2; selectedButton := bench.Operator.JoyBtnRaw; ELSE selectedX := 5000; selectedY := 5000; selectedButton := FALSE; END_IF;
joy(RawX := selectedX, RawY := selectedY, RawButton := selectedButton, Cfg := cfg, NeutralXMem := nx, NeutralYMem := ny);
IF bench.Operator.JoyBtnRaw AND NOT previousButton THEN buttonEdges := buttonEdges + 1; END_IF; previousButton := bench.Operator.JoyBtnRaw;
ADVANCE_TIME(10000000); bench.OperatorSourceActive := sourceSelected; bench(RawPosM1 := raw1, RawPosM2 := raw2);
IF sourceSelected THEN selectedX := bench.Operator.JoyXRaw_ANA1; selectedY := bench.Operator.JoyYRaw_ANA2; selectedButton := bench.Operator.JoyBtnRaw; ELSE selectedX := 5000; selectedY := 5000; selectedButton := FALSE; END_IF;
joy(RawX := selectedX, RawY := selectedY, RawButton := selectedButton, Cfg := cfg, NeutralXMem := nx, NeutralYMem := ny);
IF bench.Operator.JoyBtnRaw AND NOT previousButton THEN buttonEdges := buttonEdges + 1; END_IF; previousButton := bench.Operator.JoyBtnRaw;
ADVANCE_TIME(10000000); bench.OperatorSourceActive := sourceSelected; bench(RawPosM1 := raw1, RawPosM2 := raw2);
IF sourceSelected THEN selectedX := bench.Operator.JoyXRaw_ANA1; selectedY := bench.Operator.JoyYRaw_ANA2; selectedButton := bench.Operator.JoyBtnRaw; ELSE selectedX := 5000; selectedY := 5000; selectedButton := FALSE; END_IF;
joy(RawX := selectedX, RawY := selectedY, RawButton := selectedButton, Cfg := cfg, NeutralXMem := nx, NeutralYMem := ny);
IF bench.Operator.JoyBtnRaw AND NOT previousButton THEN buttonEdges := buttonEdges + 1; END_IF; previousButton := bench.Operator.JoyBtnRaw;
ADVANCE_TIME(10000000); bench.OperatorSourceActive := sourceSelected; bench(RawPosM1 := raw1, RawPosM2 := raw2);
IF sourceSelected THEN selectedX := bench.Operator.JoyXRaw_ANA1; selectedY := bench.Operator.JoyYRaw_ANA2; selectedButton := bench.Operator.JoyBtnRaw; ELSE selectedX := 5000; selectedY := 5000; selectedButton := FALSE; END_IF;
joy(RawX := selectedX, RawY := selectedY, RawButton := selectedButton, Cfg := cfg, NeutralXMem := nx, NeutralYMem := ny);
IF bench.Operator.JoyBtnRaw AND NOT previousButton THEN buttonEdges := buttonEdges + 1; END_IF; previousButton := bench.Operator.JoyBtnRaw;
ADVANCE_TIME(10000000); bench.OperatorSourceActive := sourceSelected; bench(RawPosM1 := raw1, RawPosM2 := raw2);
IF sourceSelected THEN selectedX := bench.Operator.JoyXRaw_ANA1; selectedY := bench.Operator.JoyYRaw_ANA2; selectedButton := bench.Operator.JoyBtnRaw; ELSE selectedX := 5000; selectedY := 5000; selectedButton := FALSE; END_IF;
joy(RawX := selectedX, RawY := selectedY, RawButton := selectedButton, Cfg := cfg, NeutralXMem := nx, NeutralYMem := ny);
IF bench.Operator.JoyBtnRaw AND NOT previousButton THEN buttonEdges := buttonEdges + 1; END_IF; previousButton := bench.Operator.JoyBtnRaw;
ADVANCE_TIME(10000000); bench.OperatorSourceActive := sourceSelected; bench(RawPosM1 := raw1, RawPosM2 := raw2);
IF sourceSelected THEN selectedX := bench.Operator.JoyXRaw_ANA1; selectedY := bench.Operator.JoyYRaw_ANA2; selectedButton := bench.Operator.JoyBtnRaw; ELSE selectedX := 5000; selectedY := 5000; selectedButton := FALSE; END_IF;
joy(RawX := selectedX, RawY := selectedY, RawButton := selectedButton, Cfg := cfg, NeutralXMem := nx, NeutralYMem := ny);
IF bench.Operator.JoyBtnRaw AND NOT previousButton THEN buttonEdges := buttonEdges + 1; END_IF; previousButton := bench.Operator.JoyBtnRaw;
ADVANCE_TIME(10000000); bench.OperatorSourceActive := sourceSelected; bench(RawPosM1 := raw1, RawPosM2 := raw2);
IF sourceSelected THEN selectedX := bench.Operator.JoyXRaw_ANA1; selectedY := bench.Operator.JoyYRaw_ANA2; selectedButton := bench.Operator.JoyBtnRaw; ELSE selectedX := 5000; selectedY := 5000; selectedButton := FALSE; END_IF;
joy(RawX := selectedX, RawY := selectedY, RawButton := selectedButton, Cfg := cfg, NeutralXMem := nx, NeutralYMem := ny);
IF bench.Operator.JoyBtnRaw AND NOT previousButton THEN buttonEdges := buttonEdges + 1; END_IF; previousButton := bench.Operator.JoyBtnRaw;
ADVANCE_TIME(10000000); bench.OperatorSourceActive := sourceSelected; bench(RawPosM1 := raw1, RawPosM2 := raw2);
IF sourceSelected THEN selectedX := bench.Operator.JoyXRaw_ANA1; selectedY := bench.Operator.JoyYRaw_ANA2; selectedButton := bench.Operator.JoyBtnRaw; ELSE selectedX := 5000; selectedY := 5000; selectedButton := FALSE; END_IF;
joy(RawX := selectedX, RawY := selectedY, RawButton := selectedButton, Cfg := cfg, NeutralXMem := nx, NeutralYMem := ny);
IF bench.Operator.JoyBtnRaw AND NOT previousButton THEN buttonEdges := buttonEdges + 1; END_IF; previousButton := bench.Operator.JoyBtnRaw;
ADVANCE_TIME(10000000); bench.OperatorSourceActive := sourceSelected; bench(RawPosM1 := raw1, RawPosM2 := raw2);
IF sourceSelected THEN selectedX := bench.Operator.JoyXRaw_ANA1; selectedY := bench.Operator.JoyYRaw_ANA2; selectedButton := bench.Operator.JoyBtnRaw; ELSE selectedX := 5000; selectedY := 5000; selectedButton := FALSE; END_IF;
joy(RawX := selectedX, RawY := selectedY, RawButton := selectedButton, Cfg := cfg, NeutralXMem := nx, NeutralYMem := ny);
IF bench.Operator.JoyBtnRaw AND NOT previousButton THEN buttonEdges := buttonEdges + 1; END_IF; previousButton := bench.Operator.JoyBtnRaw;
ASSERT_TRUE(joy.AxisCmdX.StartStop, 'Geste initial arme'); ASSERT_FALSE(selectedButton, 'Bouton armement deja relache');
sourceSelected := FALSE;
ADVANCE_TIME(10000000); bench.OperatorSourceActive := sourceSelected; bench(RawPosM1 := raw1, RawPosM2 := raw2);
IF sourceSelected THEN selectedX := bench.Operator.JoyXRaw_ANA1; selectedY := bench.Operator.JoyYRaw_ANA2; selectedButton := bench.Operator.JoyBtnRaw; ELSE selectedX := 5000; selectedY := 5000; selectedButton := FALSE; END_IF;
joy(RawX := selectedX, RawY := selectedY, RawButton := selectedButton, Cfg := cfg, NeutralXMem := nx, NeutralYMem := ny);
IF bench.Operator.JoyBtnRaw AND NOT previousButton THEN buttonEdges := buttonEdges + 1; END_IF; previousButton := bench.Operator.JoyBtnRaw;
ADVANCE_TIME(10000000); bench.OperatorSourceActive := sourceSelected; bench(RawPosM1 := raw1, RawPosM2 := raw2);
IF sourceSelected THEN selectedX := bench.Operator.JoyXRaw_ANA1; selectedY := bench.Operator.JoyYRaw_ANA2; selectedButton := bench.Operator.JoyBtnRaw; ELSE selectedX := 5000; selectedY := 5000; selectedButton := FALSE; END_IF;
joy(RawX := selectedX, RawY := selectedY, RawButton := selectedButton, Cfg := cfg, NeutralXMem := nx, NeutralYMem := ny);
IF bench.Operator.JoyBtnRaw AND NOT previousButton THEN buttonEdges := buttonEdges + 1; END_IF; previousButton := bench.Operator.JoyBtnRaw;
ADVANCE_TIME(10000000); bench.OperatorSourceActive := sourceSelected; bench(RawPosM1 := raw1, RawPosM2 := raw2);
IF sourceSelected THEN selectedX := bench.Operator.JoyXRaw_ANA1; selectedY := bench.Operator.JoyYRaw_ANA2; selectedButton := bench.Operator.JoyBtnRaw; ELSE selectedX := 5000; selectedY := 5000; selectedButton := FALSE; END_IF;
joy(RawX := selectedX, RawY := selectedY, RawButton := selectedButton, Cfg := cfg, NeutralXMem := nx, NeutralYMem := ny);
IF bench.Operator.JoyBtnRaw AND NOT previousButton THEN buttonEdges := buttonEdges + 1; END_IF; previousButton := bench.Operator.JoyBtnRaw;
ADVANCE_TIME(10000000); bench.OperatorSourceActive := sourceSelected; bench(RawPosM1 := raw1, RawPosM2 := raw2);
IF sourceSelected THEN selectedX := bench.Operator.JoyXRaw_ANA1; selectedY := bench.Operator.JoyYRaw_ANA2; selectedButton := bench.Operator.JoyBtnRaw; ELSE selectedX := 5000; selectedY := 5000; selectedButton := FALSE; END_IF;
joy(RawX := selectedX, RawY := selectedY, RawButton := selectedButton, Cfg := cfg, NeutralXMem := nx, NeutralYMem := ny);
IF bench.Operator.JoyBtnRaw AND NOT previousButton THEN buttonEdges := buttonEdges + 1; END_IF; previousButton := bench.Operator.JoyBtnRaw;
ADVANCE_TIME(10000000); bench.OperatorSourceActive := sourceSelected; bench(RawPosM1 := raw1, RawPosM2 := raw2);
IF sourceSelected THEN selectedX := bench.Operator.JoyXRaw_ANA1; selectedY := bench.Operator.JoyYRaw_ANA2; selectedButton := bench.Operator.JoyBtnRaw; ELSE selectedX := 5000; selectedY := 5000; selectedButton := FALSE; END_IF;
joy(RawX := selectedX, RawY := selectedY, RawButton := selectedButton, Cfg := cfg, NeutralXMem := nx, NeutralYMem := ny);
IF bench.Operator.JoyBtnRaw AND NOT previousButton THEN buttonEdges := buttonEdges + 1; END_IF; previousButton := bench.Operator.JoyBtnRaw;
ADVANCE_TIME(10000000); bench.OperatorSourceActive := sourceSelected; bench(RawPosM1 := raw1, RawPosM2 := raw2);
IF sourceSelected THEN selectedX := bench.Operator.JoyXRaw_ANA1; selectedY := bench.Operator.JoyYRaw_ANA2; selectedButton := bench.Operator.JoyBtnRaw; ELSE selectedX := 5000; selectedY := 5000; selectedButton := FALSE; END_IF;
joy(RawX := selectedX, RawY := selectedY, RawButton := selectedButton, Cfg := cfg, NeutralXMem := nx, NeutralYMem := ny);
IF bench.Operator.JoyBtnRaw AND NOT previousButton THEN buttonEdges := buttonEdges + 1; END_IF; previousButton := bench.Operator.JoyBtnRaw;
ADVANCE_TIME(10000000); bench.OperatorSourceActive := sourceSelected; bench(RawPosM1 := raw1, RawPosM2 := raw2);
IF sourceSelected THEN selectedX := bench.Operator.JoyXRaw_ANA1; selectedY := bench.Operator.JoyYRaw_ANA2; selectedButton := bench.Operator.JoyBtnRaw; ELSE selectedX := 5000; selectedY := 5000; selectedButton := FALSE; END_IF;
joy(RawX := selectedX, RawY := selectedY, RawButton := selectedButton, Cfg := cfg, NeutralXMem := nx, NeutralYMem := ny);
IF bench.Operator.JoyBtnRaw AND NOT previousButton THEN buttonEdges := buttonEdges + 1; END_IF; previousButton := bench.Operator.JoyBtnRaw;
ADVANCE_TIME(10000000); bench.OperatorSourceActive := sourceSelected; bench(RawPosM1 := raw1, RawPosM2 := raw2);
IF sourceSelected THEN selectedX := bench.Operator.JoyXRaw_ANA1; selectedY := bench.Operator.JoyYRaw_ANA2; selectedButton := bench.Operator.JoyBtnRaw; ELSE selectedX := 5000; selectedY := 5000; selectedButton := FALSE; END_IF;
joy(RawX := selectedX, RawY := selectedY, RawButton := selectedButton, Cfg := cfg, NeutralXMem := nx, NeutralYMem := ny);
IF bench.Operator.JoyBtnRaw AND NOT previousButton THEN buttonEdges := buttonEdges + 1; END_IF; previousButton := bench.Operator.JoyBtnRaw;
ADVANCE_TIME(10000000); bench.OperatorSourceActive := sourceSelected; bench(RawPosM1 := raw1, RawPosM2 := raw2);
IF sourceSelected THEN selectedX := bench.Operator.JoyXRaw_ANA1; selectedY := bench.Operator.JoyYRaw_ANA2; selectedButton := bench.Operator.JoyBtnRaw; ELSE selectedX := 5000; selectedY := 5000; selectedButton := FALSE; END_IF;
joy(RawX := selectedX, RawY := selectedY, RawButton := selectedButton, Cfg := cfg, NeutralXMem := nx, NeutralYMem := ny);
IF bench.Operator.JoyBtnRaw AND NOT previousButton THEN buttonEdges := buttonEdges + 1; END_IF; previousButton := bench.Operator.JoyBtnRaw;
ADVANCE_TIME(10000000); bench.OperatorSourceActive := sourceSelected; bench(RawPosM1 := raw1, RawPosM2 := raw2);
IF sourceSelected THEN selectedX := bench.Operator.JoyXRaw_ANA1; selectedY := bench.Operator.JoyYRaw_ANA2; selectedButton := bench.Operator.JoyBtnRaw; ELSE selectedX := 5000; selectedY := 5000; selectedButton := FALSE; END_IF;
joy(RawX := selectedX, RawY := selectedY, RawButton := selectedButton, Cfg := cfg, NeutralXMem := nx, NeutralYMem := ny);
IF bench.Operator.JoyBtnRaw AND NOT previousButton THEN buttonEdges := buttonEdges + 1; END_IF; previousButton := bench.Operator.JoyBtnRaw;
ASSERT_FALSE(joy.AxisCmdX.StartStop, 'Source reelle neutre selectionnee'); ASSERT_TRUE(joy.DeadmanArmed, 'Grace reelle encore active');
sourceSelected := TRUE;
ADVANCE_TIME(10000000); bench.OperatorSourceActive := sourceSelected; bench(RawPosM1 := raw1, RawPosM2 := raw2);
IF sourceSelected THEN selectedX := bench.Operator.JoyXRaw_ANA1; selectedY := bench.Operator.JoyYRaw_ANA2; selectedButton := bench.Operator.JoyBtnRaw; ELSE selectedX := 5000; selectedY := 5000; selectedButton := FALSE; END_IF;
joy(RawX := selectedX, RawY := selectedY, RawButton := selectedButton, Cfg := cfg, NeutralXMem := nx, NeutralYMem := ny);
IF bench.Operator.JoyBtnRaw AND NOT previousButton THEN buttonEdges := buttonEdges + 1; END_IF; previousButton := bench.Operator.JoyBtnRaw;
ASSERT_FALSE(joy.AxisCmdX.StartStop, 'Aucune reprise sans nouvel appui IHM a reselection simulee'); ASSERT_EQ(buttonEdges, 1, 'Aucun nouveau geste demande'); ASSERT_FALSE(selectedButton, 'Aucun nouvel appui armement');
END_TEST
